(* IEC 61131-3 sources: daoli-st-library/DL_Motion (part 9) *)

(* ---- FB_DL_AxisScrewPitchComp.st ---- *)
(*==============================================================================
 * 组件名称 (Component)  : FB_DL_AxisScrewPitchComp
 * 所属子库 (Sublibrary) : DL_Motion
 * 当前版本 (Version)    : 1.0.0
 * 兼容性   (Platform)   : CODESYS 3.5+ / TwinCAT 3 / 汇川 InoProShop / 施耐德 Machine Expert
 *                         仅依赖 Standard.library（TRUNC / ABS），零厂商私有库
 * 功能描述 (Function)   : 丝杠螺距误差分段前馈补偿：误差表 aErrTable[0..nSegCnt]
 *                         给出均匀分段节点（段长 fSegLenMm，表长 = 段数 + 1，
 *                         一致性校验）处螺距误差（mm），段内线性插值：
 *                           idx  = TRUNC(fPosMm ÷ fSegLenMm)，钳位 [0, nSegCnt−1]
 *                           fFrac = fPosMm ÷ fSegLenMm − idx，钳位 [0,1]
 *                           fCompValMm = aErrTable[idx]
 *                                        + fFrac × (aErrTable[idx+1] − aErrTable[idx])
 *                         位置先钳入表覆盖域 [0, nSegCnt×fSegLenMm]（越域置
 *                         信息码 ePosClamped），段索引防越界钳位（规格指定）；
 *                         非有限位置输出 0 并置信息码 ePosNonFin（规格指定）。
 * 接口     (Interface)  : 输入 fPosMm 轴当前位置 [mm]、aErrTable 分段误差表
 *                         （定长 0..16，[mm]）、nSegCnt 有效段数（域 [1,16]）、
 *                         fSegLenMm 每段长度（域 > 0）、bReset 复位；
 *                         输出 fCompValMm 前馈补偿值（叠加到位置设定侧）
 *                         [mm]、eErrCode 错误码、bError 故障标志。
 * 边界     (Boundary)   : ① **属主边界（写死）：本件只算螺距误差补偿量，不写
 *                         位置指令、不接管反向间隙补偿**；间隙补偿归
 *                         `FB_DL_AxisBacklashComp`。
 *                         ② 表长一致性：nSegCnt 有效段数对应节点 0..nSegCnt
 *                         共 nSegCnt+1 个，超出定长 17（nSegCnt > 16）或
 *                         nSegCnt < 1 → 锁存故障（表长=段数+1 一致性校验，
 *                         规格指定），冻结输出 0。
 *                         ③ 位置域钳位：fPosMm < 0 钳 0、> nSegCnt×fSegLenMm
 *                         钳上界，置信息码 ePosClamped（量值方向可饱和）。
 *                         ④ 非有限判据（R79 双判）先行于一切换算：非有限时
 *                         输出 0、信息码 ePosNonFin，不污染插值。
 *                         ⑤ 组态闸：fSegLenMm <= 0 → 锁存故障（除数前置闸，
 *                         结构性无除零），冻结输出 0，解除沿 = bReset 上升沿。
 *                         ⑥ TRUNC 取整前位置已过非有限闸与域钳位（无溢出
 *                         取整路径）。
 *                         ⑦ 零全局耦合（无 GVL / VAR_EXTERNAL / 物理地址）。
 * 分工声明 (Scope)      : 与 `FB_DL_AxisBacklashComp` 分工：反向间隙（双区滞回）
 *                         归那件、螺距分段误差（单值表）归本件；与
 *                         `FB_DL_CamTableInterp` 分工：凸轮表插值归那件。
 * 来源标签 (Source Tag) : 自研线（分段线性插值为公开数值方法 clean-room）
 * 码表     (Codes)      : 本件不占用任何全局数字码位。出口为 LREAL 补偿值 +
 *                         ENUM 错误码；数字码位待主控收口阶段统一派号。
 * 红线自检 (Redline)    : R1 ✓ 零 GVL/VAR_EXTERNAL ｜ R2 ✓ 零 %I/%Q/%M ｜ R3 ✓ 纯 IEC 61131-3
 *                         R4 ✓ 索引钳位 + 表长一致性 + 除数前置闸 + 非有限先行
 *                         ｜ R5 ✓ 声明逐行同行双语注释
 *                         R6 N/A（无 ENUM 状态机） ｜ R7 ✓ 一 R_TRIG 段 0 无条件刷新
 * 修订历史 (Revision)   : 2026-11-20  v1.0.0  R50 首版（批次 2 · 序号 7）
 * 验收向量 (Acceptance) : ① fSegLenMm=10, nSegCnt=2, aErrTable=[0.0, 0.01, 0.03]
 *                         （mm）：fPosMm=5 → 段 0 半程 → 0.0 + 0.5×0.01 =
 *                         0.005 mm；fPosMm=15 → 段 1 半程 → 0.01 + 0.5×0.02
 *                         = 0.02 mm，均 eOk；② fPosMm=25 → 钳上界 20 → 段 1
 *                         终点 → 0.03 mm，ePosClamped；③ nSegCnt=0 → 锁存
 *                         eCfgBad，输出 0；④ fPosMm=NaN → 输出 0，
 *                         ePosNonFin。
 *==============================================================================*)

(*-----------------------------------------------------------------------------
 * 枚举: E_DL_SpcErr（错误码；信息级不置 bError，故障级恒伴 bError=TRUE）
 *----------------------------------------------------------------------------*)
TYPE E_DL_SpcErr :
(
    eOk         := 0,   // 正常 / Normal
    eCfgBad     := 1,   // 故障级：段数/段长组态非法（表长=段数+1 破坏） / Fault: segment config illegal
    ePosClamped := 2,   // 信息级：位置越表域已钳位 / Info: position clamped into table domain
    ePosNonFin  := 3    // 信息级：位置非有限，输出 0 / Info: position non-finite, output zero
);
END_TYPE

FUNCTION_BLOCK FB_DL_AxisScrewPitchComp
VAR_INPUT
    fPosMm    : LREAL := 0.0;                  // 轴当前位置 [mm] / Axis present position [mm]
    aErrTable : ARRAY[0..16] OF LREAL;         // 分段误差表（节点 0..nSegCnt） [mm] / Segmented error table [mm]
    nSegCnt   : UDINT := 8;                    // 有效段数（表长 = 段数+1），域 [1,16] [段] / Valid segment count
    fSegLenMm : LREAL := 10.0;                 // 每段长度，域 > 0 [mm] / Segment length [mm]
    bReset    : BOOL := FALSE;                 // 复位，上升沿清组态故障锁存 [-] / Reset, rising edge clears cfg latch
END_VAR
VAR_OUTPUT
    fCompValMm : LREAL;                        // 前馈补偿值（叠加位置设定侧） [mm] / Feedforward compensation [mm]
    eErrCode   : E_DL_SpcErr;                  // 错误码出口 / Error code outlet
    bError     : BOOL;                         // 故障标志（组态锁存） [-] / Error flag, latched
END_VAR
VAR
    _nIdx     : DINT;                          // 段索引（钳位后，域 [0, nSegCnt−1]） [-] / Clamped segment index
    _fScaled  : LREAL;                         // 位置按段长标度值（无量纲段数） [段] / Position scaled by segment length
    _fFrac    : LREAL;                         // 段内分数（钳位 [0,1]） [-] / In-segment fraction
    _fPosUse  : LREAL;                         // 钳入表域后的位置 [mm] / Position clamped into domain
    _fPosMax  : LREAL;                         // 表覆盖域上界 = nSegCnt×fSegLenMm [mm] / Table domain ceiling
    _bNonFin  : BOOL;                          // 位置非有限当拍量 [-] / Position non-finite this scan
    _bClamped : BOOL;                          // 本拍发生位置钳位 [-] / Position clamped this scan
    _bCfgBad  : BOOL;                          // 组态非法当拍量 [-] / Illegal configuration this scan
    _bErrLatch: BOOL;                          // 组态故障锁存位（解除沿 = bReset 上升沿） / Latched config fault
    rtReset   : R_TRIG;                        // 复位沿实例，段 0 无条件调用 / Reset edge instance
END_VAR
VAR CONSTANT
    DL_SPC_NMAX  : DINT := 16;                 // 段数上限（表定长 0..16 共 17 节点） [段] / Segment count ceiling
    DL_SPC_NMIN  : DINT := 1;                  // 段数下限 [段] / Segment count floor
    DL_SPC_ZERO  : LREAL := 0.0;               // 域下界与判零基准 [mm] / Domain floor and zero base
    DL_SPC_ONE   : LREAL := 1.0;               // 分数钳位上界 [-] / Fraction ceiling
END_VAR

(* —— 段 0：非有限判 + 组态闸 + 沿刷新 —— *)
_bNonFin := (fPosMm <> fPosMm) OR ((fPosMm - fPosMm) <> DL_SPC_ZERO);   // 位置非有限（R79 双判） / Position non-finite
_bCfgBad := (fSegLenMm <= DL_SPC_ZERO);        // 段长域闸（除数前置） / Segment length gate
IF (UDINT_TO_DINT(nSegCnt) < DL_SPC_NMIN) OR (UDINT_TO_DINT(nSegCnt) > DL_SPC_NMAX) THEN
    _bCfgBad := TRUE;                          // 表长=段数+1 一致性破坏（规格②） / Table length consistency violated
END_IF
rtReset(CLK := bReset);                        // 复位沿，每拍必调 / Reset edge, every scan

(* —— 段 1：复位沿与组态锁存 —— *)
IF rtReset.Q THEN
    _bErrLatch := FALSE;                       // 清组态锁存（R188 声明：解除沿 = bReset 上升沿） / Clear cfg latch
END_IF
IF _bCfgBad AND (NOT _bErrLatch) THEN
    _bErrLatch := TRUE;                        // 锁存 / Latch
END_IF

(* —— 段 2：位置域钳位（故障期跳过；非有限跳过） —— *)
_bClamped := FALSE;                            // 钳位量预清 / Clamp preset
_fPosUse := DL_SPC_ZERO;                       // 安全侧起步 0 / Safe-side start zero
_fPosMax := UDINT_TO_LREAL(nSegCnt) * fSegLenMm;   // 表域上界 [mm] / Domain ceiling
IF (NOT _bErrLatch) AND (NOT _bNonFin) THEN
    _fPosUse := fPosMm;                        // 位置工作副本 / Position working copy
    IF _fPosUse < DL_SPC_ZERO THEN
        _fPosUse := DL_SPC_ZERO;               // 下越域钳 0 / Clamp low to zero
        _bClamped := TRUE;                     // 记钳位 / Mark clamp
    ELSIF _fPosUse > _fPosMax THEN
        _fPosUse := _fPosMax;                  // 上越域钳上界 / Clamp high to ceiling
        _bClamped := TRUE;                     // 记钳位 / Mark clamp
    END_IF
END_IF

(* —— 段 3：分段线性插值（索引与分数双重钳位，防越界） —— *)
IF (NOT _bErrLatch) AND (NOT _bNonFin) THEN
    _fScaled := _fPosUse / fSegLenMm;          // 标度值（除数已过闸，结构性无除零） / Scaled value
    _nIdx := LREAL_TO_DINT(TRUNC(_fScaled));   // 段索引取整（域已钳，无溢出） / Segment index by TRUNC
    IF _nIdx > (UDINT_TO_DINT(nSegCnt) - 1) THEN
        _nIdx := UDINT_TO_DINT(nSegCnt) - 1;   // 索引上钳（规格：防越界钳位） / Clamp index high
    END_IF
    IF _nIdx < 0 THEN
        _nIdx := 0;                            // 索引下钳 / Clamp index low
    END_IF
    _fFrac := _fScaled - DINT_TO_LREAL(_nIdx);   // 段内分数（索引升位实数化） / In-segment fraction
    IF _fFrac < DL_SPC_ZERO THEN
        _fFrac := DL_SPC_ZERO;                 // 分数下钳 / Clamp fraction low
    END_IF
    IF _fFrac > DL_SPC_ONE THEN
        _fFrac := DL_SPC_ONE;                  // 分数上钳 / Clamp fraction high
    END_IF
    fCompValMm := aErrTable[_nIdx] + _fFrac * (aErrTable[_nIdx + 1] - aErrTable[_nIdx]);   // 段内线性插值（_nIdx+1 <= nSegCnt 表内） / Linear interpolation
ELSE
    fCompValMm := DL_SPC_ZERO;                 // 故障/非有限安全侧输出 0（规格④） / Safe-side zero output
END_IF

(* —— 段 4：出口单点映射（错误码归约，R191） —— *)
IF _bErrLatch THEN
    bError := TRUE;                            // 故障标志（R45 配对） / Error flag
    eErrCode := E_DL_SpcErr.eCfgBad;           // 故障级码 / Fault code
ELSE
    bError := FALSE;                           // 无故障级条件 / No fault
    IF _bNonFin THEN
        eErrCode := E_DL_SpcErr.ePosNonFin;    // 信息级：非有限口径 / Info: non-finite
    ELSIF _bClamped THEN
        eErrCode := E_DL_SpcErr.ePosClamped;   // 信息级：越域钳位口径 / Info: clamped
    ELSE
        eErrCode := E_DL_SpcErr.eOk;           // 正常 / Normal
    END_IF
END_IF

END_FUNCTION_BLOCK

(* ---- FB_DL_AxisSoftLimitGuard.st ---- *)
(*
    FB_DL_AxisSoftLimitGuard —— 轴软限位守卫（位置 + 速度前馈预判减速请求）
    ------------------------------------------------------------------
    组件名称  : FB_DL_AxisSoftLimitGuard
    分类      : DL_Motion / LimitGuard
    前缀      : FB_DL_
    版本      : 1.0.0
    溯源      : 借鉴点 —— 运动控制领域「软限位 + 提前减速（预判停距）」的通行语义：
                仅用位置比较只能撞限位后才发现（已超程），故必须用当前速度按
                允许减速度反算停距，把「当前位置 + 本周期位移 + 停距」作为预判
                可达位置，与限位比较后提前发出减速请求；越限后锁存并禁止该方向
                运动（方向互锁）。该语义与 PLCopen Motion Control 公开规范中
                「软限位监视 / 方向禁止」的功能描述一致。
                clean-room 声明 —— 零代码行复制；本件不含任何厂商运动指令
                （不调用 MC_* 功能块、不使用任何厂商专有数据类型），停距预判、
                方向互锁、闸门、码位与双语文档全部自有。
                许可证 —— 本件 MIT；来源标签 s7motion 仅指该语义在公开厂商文档
                中的功能描述，文档不属代码，无许可继承。
    平台      : 纯 IEC 61131-3，CODESYS 3.5 / TwinCAT 3 / InoProShop / Machine Expert 通用
    作者      : 道莅代码库 · PLC编程专家（R70 构建轮 · 批 3 · N8）
    ------------------------------------------------------------------
    功能说明  : 预判模型（逐项写清，便于现场复核）：
                  fSpan := ABS(fVel) * fScanSec               本周期位移（速度前馈项，[mm]）
                  fStop := fVel * fVel / (2 * fDecel)         停距（等减速度制动距离，[mm]）
                  fPred := fPos + fVel * fScanSec + 符号(fVel) * fStop   预判可达位置 [mm]
                判据：
                  正向减速请求 bDecelPos := fVel > 0 且 fPred > (fPosMax - fMargin)
                  负向减速请求 bDecelNeg := fVel < 0 且 fPred < (fPosMin + fMargin)
                  正向禁止 bInhibitPos := 越限锁存 或 fPos >= fPosMax
                  负向禁止 bInhibitNeg := 越限锁存 或 fPos <= fPosMin
                除法面（唯一除法）：除子为 (2 * fDecel)，进入除法前经**两道结构闸**
                校验 fDecel > 0 与 (2 * fDecel) > 0，两者同时成立才落除法；
                闸不成立时整个预判段被跳过（不落除法、不发减速请求、不写
                fPredPos），并由组态闸在段 4 置 0501 锁存。
                其余算式一律用乘加（余量比较改写为 fMargin * 2 >= 行程），
                故本件全部代码中只有一个除法点。
                越限锁存：fPos 越过任一限位即锁存 0503，bReset 上升沿解除；
                锁存期内两个禁止方向位**恒为 TRUE**（双方向全禁，因为越限后
                任何方向都可能加剧超程，需人工确认后复位）。
    错误码    : 16#0002_0501 组态非法（限位反置 / 减速度非正 / 回退余量为负 / 非有限），锁存 —— 故障级
                16#0002_0502 位置或速度非有限，锁存 —— 故障级
                16#0002_0503 越限（位置越过软限位），锁存 —— 故障级
    码位总账  : 0501 / 0502 / 0503 用（均故障级）；无信息级码（减速请求与禁止位已可观测）
    状态机    : N/A —— 无顺序相（逐拍组合判据 + 越限锁存），无 ENUM / CASE
    边界与披露: 一 组态闸（R272 逐项点名）：fPosMax > fPosMin；fDecel > 0；
                   fMargin >= 0 且 fMargin < (fPosMax - fPosMin) / 2（余量不得吞没
                   整个行程）；fScanSec > 0；上述量与 fPos / fVel 全部纳入
                   NaN 自反判 + Inf 差值自反判 + 幅值 1E9 上界筛查；
                二 定时器 / 沿实例：仅 _rtReset 一个沿实例，在段 2 无条件调用；
                   本件不含 TON / TOF / TP，故无定时器跳过风险；
                三 出口语义（R191）：bDecelPos / bDecelNeg 为**逐拍重算**的请求位，
                   bInhibitPos / bInhibitNeg 为组合位（越限锁存 或 位置到限），
                   bBeyond 为越限锁存镜像；三者名实同源、无混用；
                四 失能（bEn = FALSE）：减速请求清零、禁止位**保持有效**
                   （安全方向：失能不得放开方向禁止），bBusy 清零，锁存位不被清除；
                五 本件不做任何运动指令下发，只输出布尔许可 / 请求位，由上层
                   运动层转换为 MC_Halt / 减速倍率等动作 —— 保持硬件与厂商无关；
                六 零全局变量、零 VAR_EXTERNAL、零物理地址、零数组下标。
    修订记录  : 2026-11-22 v1.0.0 首次入库（R70 构建轮 · 批 3 · N8）
*)
FUNCTION_BLOCK FB_DL_AxisSoftLimitGuard
VAR_INPUT
    bEn       : BOOL := TRUE;              (* 使能，[标志] / the enable *)
    bReset    : BOOL := FALSE;             (* 越限复位（上升沿有效），[标志] / the overrun reset, rising edge *)
    fPos      : LREAL := 0.0;              (* 轴当前位置（编码器反馈），[mm] / the axis position feedback *)
    fVel      : LREAL := 0.0;              (* 轴当前速度（反馈或指令前馈），[mm/s] / the axis velocity *)
    fPosMax   : LREAL := 1000.0;           (* 正向软限位，[mm]，须 > fPosMin / the positive soft limit *)
    fPosMin   : LREAL := 0.0;              (* 负向软限位，[mm]，须 < fPosMax / the negative soft limit *)
    fDecel    : LREAL := 1000.0;           (* 允许减速度幅值，[mm/s^2]，须 > 0 / the allowed deceleration magnitude *)
    fScanSec  : LREAL := 0.004;            (* 任务周期折算秒数，[s]，须 > 0 / the task period in seconds *)
    fMargin   : LREAL := 20.0;             (* 提前减速余量，[mm]，须 >= 0 / the early deceleration margin *)
END_VAR
VAR_OUTPUT
    bDecelPos   : BOOL;                    (* 正向减速请求，[标志] / the positive direction deceleration request *)
    bDecelNeg   : BOOL;                    (* 负向减速请求，[标志] / the negative direction deceleration request *)
    bInhibitPos : BOOL;                    (* 正向运动禁止，[标志] / the positive direction inhibited *)
    bInhibitNeg : BOOL;                    (* 负向运动禁止，[标志] / the negative direction inhibited *)
    bBeyond     : BOOL;                    (* 越限锁存镜像，[标志] / the overrun latch image *)
    fPredPos    : LREAL;                   (* 预判可达位置（供诊断），[mm] / the predicted reachable position *)
    bBusy       : BOOL;                    (* 减速请求有效（占用中），[标志] / a deceleration request is active *)
    bValid      : BOOL;                    (* 出口可信（无锁存故障），[标志] / the outlets are trustworthy *)
    bError      : BOOL;                    (* 故障标志，锁存故障时为 TRUE / the fault flag, raised while latched *)
    nErrCode    : UDINT;                   (* 错误码，0 = 正常，锁存回放 / the error id, 0 = ok, replayed *)
END_VAR
VAR
    _rtReset    : R_TRIG;                  (* 复位上升沿实例（无条件调用）/ the reset rising edge instance *)
    _bFault     : BOOL;                    (* 组态 / 输入故障锁存位 / the configuration and input fault latch *)
    _bBeyond    : BOOL;                    (* 越限保持量，仅 bReset 上升沿解除 / the overrun hold *)
    _nCodeLatch : UDINT;                   (* 故障锁存码（0501 / 0502 / 0503）/ the fault code latch *)
    _bCfgBad    : BOOL;                    (* 组态非法标志（逐拍重算）/ the configuration fault flag *)
    _bInBad     : BOOL;                    (* 位置或速度非有限标志（逐拍重算）/ the input fault flag *)
    _fSpan      : LREAL;                   (* 本周期位移，[mm] / the travel within one period *)
    _fStop      : LREAL;                   (* 制动停距，[mm] / the braking distance *)
    _fPred      : LREAL;                   (* 预判可达位置（内部），[mm] / the predicted reachable position, internal *)
    _fSign      : LREAL;                   (* 速度符号的实数形式（1.0 / 0.0 / -1.0），[无量纲] / the velocity sign as a real *)
END_VAR
VAR CONSTANT
    DL_ASG_FMAX : LREAL := 1.0E9;          (* 非有限筛查幅值上限，[工程单位] / the finiteness screening cap *)
END_VAR

// 段 1｜出口预置（R256 统一出口预置）/ segment 1, preset every outlet
bDecelPos   := FALSE;                      // 正向减速请求预清零 / preset the positive request false
bDecelNeg   := FALSE;                      // 负向减速请求预清零 / preset the negative request false
bInhibitPos := FALSE;                      // 正向禁止预清零（段 7 按安全方向重算）/ preset the positive inhibit false
bInhibitNeg := FALSE;                      // 负向禁止预清零 / preset the negative inhibit false
bBeyond     := FALSE;                      // 越限镜像预清零 / preset the overrun image false
fPredPos    := 0.0;                        // 预判位置预置零 / preset the predicted position
bBusy       := FALSE;                      // 忙碌标志预清零 / preset the busy flag false
bValid      := FALSE;                      // 可用标志预置假，健康路径再置真 / preset valid false
bError      := FALSE;                      // 故障标志预清零 / preset the error flag false
nErrCode    := 0;                          // 错误码预置无错 / preset the code to zero
_fSign      := 0.0;                        // 速度符号预置零 / preset the sign to zero

// 段 2｜沿实例无条件调用（规则 ⑦，本件无 TON / TOF / TP）/ segment 2, the reset edge instance
_rtReset(CLK := bReset);                   // 复位沿，每周期无条件刷新 / the reset edge, refreshed every scan

// 段 3｜越限解除：唯一可到达的清除边（R188）/ segment 3, the only overrun release edge
IF _rtReset.Q THEN                         // 复位上升沿 / the reset rising edge
    _bBeyond := FALSE;                     // 解除越限保持 / release the overrun hold
    IF _nCodeLatch = 16#0002_0503 THEN     // 锁存码为越限时才清码（组态 / 输入码保持到修复）/ clear the code only when it was the overrun
        _nCodeLatch := 0;                  // 清锁存码 / clear the latched code
    END_IF
END_IF

// 段 4｜组态守卫（R272 逐项点名）/ segment 4, the configuration guard
_bCfgBad := (fPosMax <= fPosMin)                                     // 限位反置或重合 / the limits reversed or coincident
         OR (fDecel <= 0.0)                                          // 减速度非正（除子域非法）/ a non positive deceleration
         OR (fScanSec <= 0.0)                                        // 任务周期非正 / a non positive task period
         OR (fMargin < 0.0)                                          // 余量为负 / a negative margin
         OR (fMargin * 2.0 >= (fPosMax - fPosMin))                   // 余量吞没行程（改用乘 2，本式不落除法）/ the margin swallows the stroke, no division here
         OR (fPosMax <> fPosMax) OR ((fPosMax - fPosMax) <> 0.0) OR (ABS(fPosMax) > DL_ASG_FMAX)
         OR (fPosMin <> fPosMin) OR ((fPosMin - fPosMin) <> 0.0) OR (ABS(fPosMin) > DL_ASG_FMAX)
         OR (fDecel <> fDecel) OR ((fDecel - fDecel) <> 0.0) OR (ABS(fDecel) > DL_ASG_FMAX)
         OR (fScanSec <> fScanSec) OR ((fScanSec - fScanSec) <> 0.0) OR (ABS(fScanSec) > DL_ASG_FMAX)
         OR (fMargin <> fMargin) OR ((fMargin - fMargin) <> 0.0) OR (ABS(fMargin) > DL_ASG_FMAX);

// 段 5｜输入守卫：位置与速度非有限 / segment 5, the position and velocity guard
_bInBad := (fPos <> fPos) OR ((fPos - fPos) <> 0.0) OR (ABS(fPos) > (DL_ASG_FMAX * 10.0))
        OR (fVel <> fVel) OR ((fVel - fVel) <> 0.0) OR (ABS(fVel) > (DL_ASG_FMAX * 10.0));

// 段 6｜首次成因锁存（故障期不重推断，R189）/ segment 6, the first cause latch
IF NOT _bFault THEN                        // 未锁存才登记 / register only while healthy
    IF _bCfgBad THEN                       // 组态非法优先 / the configuration first
        _bFault     := TRUE;               // 置锁存 / latch it
        _nCodeLatch := 16#0002_0501;       // 故障级：组态非法 / fault level: an illegal configuration
    ELSIF _bInBad THEN                     // 输入非有限 / an input is non finite
        _bFault     := TRUE;               // 置锁存 / latch it
        _nCodeLatch := 16#0002_0502;       // 故障级：输入非有限 / fault level: an input is non finite
    END_IF
END_IF

// 段 7｜越限判定与方向禁止（安全方向：越限后双向全禁）/ segment 7, the overrun verdict and the direction inhibits
IF bEn AND NOT _bFault THEN                // 使能与无故障才判越限 / judge the overrun only while enabled and healthy
    IF (fPos > fPosMax) OR (fPos < fPosMin) THEN   // 位置越过任一软限位 / the position passed a soft limit
        IF NOT _bBeyond THEN               // 首次越限才登记码（不重推断）/ register the code once
            _bBeyond    := TRUE;           // 置越限保持 / hold the overrun
            _nCodeLatch := 16#0002_0503;   // 故障级：越限 / fault level: an overrun
        END_IF
    END_IF
    bInhibitPos := _bBeyond OR (fPos >= fPosMax);  // 正向禁止：越限锁存 或 位置到正限 / the positive inhibit
    bInhibitNeg := _bBeyond OR (fPos <= fPosMin);  // 负向禁止：越限锁存 或 位置到负限 / the negative inhibit
ELSE                                       // 失能或故障：禁止位保持安全侧（不放开）/ disabled or faulted, keep the inhibits safe
    bInhibitPos := TRUE;                   // 正向保持禁止 / keep the positive direction inhibited
    bInhibitNeg := TRUE;                   // 负向保持禁止 / keep the negative direction inhibited
END_IF

// 段 8｜预判停距与减速请求（唯一除法，除子先经结构闸）/ segment 8, the predictive request
IF bEn AND NOT _bFault AND NOT _bBeyond THEN   // 健康且未越限才做预判 / predict only while healthy and inside the limits
    IF fDecel > 0.0 THEN                       // 结构闸一：减速度为正 / gate one, the deceleration is positive
        IF (2.0 * fDecel) > 0.0 THEN           // 结构闸二：除子为正（禁除零，规则 ④）/ gate two, the divisor is positive
            _fSpan := ABS(fVel) * fScanSec;    // 本周期位移（速度前馈项）/ the travel within one period
            _fStop := (fVel * fVel) / (2.0 * fDecel); // 制动停距（唯一除法）/ the braking distance, the only division
            IF fVel > 0.0 THEN                 // 正向运动 / moving in the positive direction
                _fSign := 1.0;                 // 符号为正 / the sign is positive
            ELSIF fVel < 0.0 THEN              // 负向运动 / moving in the negative direction
                _fSign := -1.0;                // 符号为负 / the sign is negative
            ELSE                               // 静止 / at standstill
                _fSign := 0.0;                 // 符号为零（停距不计方向）/ the sign is zero
            END_IF
            _fPred := fPos + (fVel * fScanSec) + (_fSign * _fStop); // 预判可达位置 / the predicted reachable position
            fPredPos := _fPred;                // 预判位置出口（诊断用）/ the predicted position outlet
            bDecelPos := (fVel > 0.0) AND (_fPred > (fPosMax - fMargin));  // 正向提前减速请求 / the positive early request
            bDecelNeg := (fVel < 0.0) AND (_fPred < (fPosMin + fMargin));  // 负向提前减速请求 / the negative early request
        END_IF
    END_IF
END_IF

// 段 9｜出口映射（名实双出口同源，R191）/ segment 9, the outlet mapping
bBeyond  := _bBeyond;                      // 越限镜像 = 保持量 / the overrun image mirrors the hold
bBusy    := bDecelPos OR bDecelNeg;        // 减速请求有效即占用 / a request is active
bError   := _bFault OR _bBeyond;           // 故障标志 = 锁存故障 或 越限 / the fault flag, the latch or the overrun
bValid   := bEn AND NOT bError;            // 出口可信条件 / the outlets are trustworthy
IF _bBeyond THEN                           // 越限优先归因 / the overrun takes precedence
    nErrCode := 16#0002_0503;              // 故障级：越限 / fault level: an overrun
ELSE                                       // 非越限 / no overrun
    nErrCode := _nCodeLatch;               // 回放锁存码 / replay the latched code
END_IF
END_FUNCTION_BLOCK

(* ---- FB_DL_AxisSoftLimitPredict.st ---- *)
(*
  Name        : FB_DL_AxisSoftLimitPredict
  Category    : DL_Motion
  Version     : 1.0.0
  Purpose     : 软限位超程预测：按当前速度与最大减速度预算停车距离 s = v²/(2a)，与到限位余量比较，提前发出减速请求（预测式，非反应式拦截）；/ Predict soft-limit overtravel: budget the stopping distance s = v^2/(2a) from current velocity and maximum deceleration, compare with the remaining margin and raise a deceleration request in advance
  溯源        : 借 t2-4-s7-motion 的分类/参数域组织，clean-room 实现
  Boundary    : ① 组态闸：最大减速度 <= eps / 余量 <= 0 / 上限须大于下限 / 扫描周期 <= 0 → 锁存故障；
                ② 除子闸：2a 在组态闸后使用（a > eps 已保证）；v² 为乘性无除法；
                ③ 仅对「朝限位运动」的方向预测：速度为 0 时不请求减速（无预测语义）；
                ④ 输出为「请求」，不直接写速度/位置（属主边界：执行由运动控制层完成）；
                ⑤ 所有比较用容差或直比，禁浮点等值比较。
*)
TYPE E_DL_AslpState :
(
    eIdle  := 0,                             (* 未使能 / Disabled *)
    ePred  := 10,                            (* 预测运行 / Predicting *)
    eFault := 90                             (* 故障锁存相 / Fault latched *)
);
END_TYPE

TYPE E_DL_AslpCause :
(
    eNone       := 0,                        (* 无故障成因 / No cause *)
    eCfgIllegal := 1,                        (* 组态非法：减速度/余量/限位越域 / Illegal config *)
    ePhaseBad   := 2                         (* 非法相位兜底 / Illegal phase fallback *)
);
END_TYPE

FUNCTION_BLOCK FB_DL_AxisSoftLimitPredict
VAR_INPUT
    fPosNow   : REAL := 0.0;                 (* 当前实际位置 [mm] / Current position *)
    fVelNow   : REAL := 0.0;                 (* 当前速度（带符号）[mm/s] / Current velocity, signed *)
    fDecMax   : REAL := 5000.0;              (* 最大可用减速度，域 > 0 [mm/s²] / Maximum deceleration, > 0 *)
    fLimPos   : REAL := 1000.0;              (* 正向软限位 [mm] / Positive soft limit *)
    fLimNeg   : REAL := -1000.0;             (* 负向软限位 [mm] / Negative soft limit *)
    fMargin   : REAL := 5.0;                 (* 提前量（在停车距离上附加），域 >= 0 [mm] / Lead margin, >= 0 *)
    bEnable   : BOOL := TRUE;                (* 预测使能 [-] / Enable *)
    bReset    : BOOL := FALSE;               (* 复位命令，上升沿清输出与故障 [-] / Reset command *)
END_VAR
VAR_OUTPUT
    fStopDist : REAL;                        (* 停车距离预算 v²/(2a) [mm] / Budgeted stopping distance *)
    fDistPos  : REAL;                        (* 到正向限位的余量 [mm] / Remaining distance to positive limit *)
    fDistNeg  : REAL;                        (* 到负向限位的余量 [mm] / Remaining distance to negative limit *)
    bDecelReq : BOOL;                        (* 减速请求（预算 + 余量 >= 可用余量）[-] / Deceleration request *)
    bOvershoot: BOOL;                        (* 已判定越界（余量 <= 提前量）[-] / Already out of margin *)
    nDir      : INT;                         (* 运动方向：+1 正 / -1 负 / 0 停 [-] / Motion direction *)
    eState    : E_DL_AslpState;              (* 状态出口 / State outlet *)
    eCause    : E_DL_AslpCause;              (* 故障成因出口（R190 归因唯一） / Fault cause outlet *)
    bError    : BOOL;                        (* 故障锁存标志 [-] / Fault latch flag *)
END_VAR
VAR
    _eState  : E_DL_AslpState := E_DL_AslpState.eIdle;   (* 内部相位（CASE 唯一写入目标） / Internal phase *)
    _eCause  : E_DL_AslpCause := E_DL_AslpCause.eNone;   (* 故障成因锁存量 / Latched cause *)
    rtReset  : R_TRIG;                       (* 复位沿实例，段 0 无条件调用 / Reset edge instance *)
    _bFault  : BOOL;                         (* 故障锁存位 / Latched fault bit *)
    _bCfgBad : BOOL;                         (* 组态非法当拍量 / Illegal config this scan *)
    _bFinite : BOOL;                         (* 输入有限性当拍量 / Input finiteness *)
    _fStop   : REAL;                         (* 停车距离中间量 [mm] / Stopping distance intermediate *)
    _fNeed   : REAL;                         (* 预算 + 提前量（总需距）[mm] / Required distance *)
    _fAbsVel : REAL;                         (* 速度绝对値（距离预算用）[mm/s] / Absolute velocity *)
    _nDir    : INT;                          (* 方向判定中间量 [-] / Direction intermediate *)
    _fZero   : REAL;                         (* 实数零常量 [-] / Real zero constant *)
END_VAR
VAR CONSTANT
    DL_ASLP_EPS : REAL := 1.0E-6;            (* 判零容差（速度/减速度）[mm/s] / Epsilon *)
    DL_ASLP_TWO : REAL := 2.0;               (* 停车距离公式常量 2 [-] / Formula constant *)
    DL_ASLP_DIRP: INT  := 1;                 (* 正方向编码 [-] / Positive direction code *)
    DL_ASLP_DIRN: INT  := -1;                (* 负方向编码 [-] / Negative direction code *)
    DL_ASLP_DIR0: INT  := 0;                 (* 静止编码 [-] / Standstill code *)
END_VAR

(* —— 段 0：当拍判据派生 + 实例无条件刷新（R228A） —— *)
_bCfgBad := (fDecMax <= DL_ASLP_EPS)                                           (* 减速度正域闸（除零前置） / Deceleration gate *)
            OR (fMargin < 0.0)                                                 (* 提前量非负闸 / Margin gate *)
            OR ((fLimPos - fLimNeg) <= DL_ASLP_EPS);                           (* 限位区间正域闸 / Limit span gate *)
rtReset(CLK := bReset);                                                        (* 复位沿每拍必调 / Reset edge every scan *)
_bFinite := (fPosNow = fPosNow) AND (fVelNow = fVelNow)                        (* NaN 自反闸 / NaN reflex gates *)
            AND ((fPosNow - fPosNow) = (fPosNow - fPosNow))                    (* 位置 Inf 闸 / Position Inf gate *)
            AND ((fVelNow - fVelNow) = (fVelNow - fVelNow));                   (* 速度 Inf 闸 / Velocity Inf gate *)
_fZero := 0.0;                                                                 (* 零常量装载 / Zero constant load *)

(* —— 段 1：单拍量预清零（R107） —— *)
bDecelReq := FALSE;                                                            (* 减速请求预清 / Request preset *)
bOvershoot := FALSE;                                                           (* 越界判据预清 / Overshoot preset *)
nDir := DL_ASLP_DIR0;                                                          (* 方向出口预清为静止 / Direction preset *)
fStopDist := 0.0;                                                              (* 停车距离预清 / Stop distance preset *)

(* —— 段 2：复位沿处理（作用域：清故障 + 清输出 + 迁 eIdle，R283 逐项声明） —— *)
IF rtReset.Q THEN
    _bFault := FALSE;                                                          (* 清故障锁存 / Clear fault *)
    _eCause := E_DL_AslpCause.eNone;                                           (* 清成因 / Clear cause *)
    fStopDist := 0.0;                                                          (* 清距离预算出口 / Clear budget outlet *)
    fDistPos := 0.0;                                                           (* 清正向余量出口 / Clear positive margin *)
    fDistNeg := 0.0;                                                           (* 清负向余量出口 / Clear negative margin *)
    bDecelReq := FALSE;                                                        (* 清减速请求 / Clear request *)
    bOvershoot := FALSE;                                                       (* 清越界判据 / Clear overshoot *)
    nDir := DL_ASLP_DIR0;                                                      (* 方向回静止 / Direction to standstill *)
    _eState := E_DL_AslpState.eIdle;                                           (* 迁未使能相 / Back to idle *)
END_IF

(* —— 段 3：组态故障锁存（锁存至复位沿，R189） —— *)
IF _bCfgBad AND NOT _bFault THEN
    _bFault := TRUE;                                                           (* 锁存故障位 / Latch fault *)
    _eCause := E_DL_AslpCause.eCfgIllegal;                                     (* 成因：组态非法 / Cause: illegal config *)
    _eState := E_DL_AslpState.eFault;                                          (* 同步迁故障相 / Migrate to fault *)
END_IF

(* —— 段 4：CASE 主状态机（ELSE 兜底迁 eFault，红线 6） —— *)
CASE _eState OF
    E_DL_AslpState.eIdle:                                                      (* 未使能：不预测 / Disabled *)
        fDistPos := fLimPos - fPosNow;                                         (* 正向余量仍实时镜像（只读观测） / Positive margin mirror *)
        fDistNeg := fPosNow - fLimNeg;                                         (* 负向余量镜像 / Negative margin mirror *)
        IF bEnable AND NOT _bFault THEN
            _eState := E_DL_AslpState.ePred;                                   (* 使能进入预测 / Enter predicting *)
        END_IF
    E_DL_AslpState.ePred:                                                      (* 预测相：停车距离预算 + 双侧余量判据 / Predicting *)
        IF NOT bEnable THEN
            _eState := E_DL_AslpState.eIdle;                                   (* 失能回未使能 / Back to idle *)
        ELSIF _bFinite THEN
            fDistPos := fLimPos - fPosNow;                                     (* 到正向限位余量（可负 = 已越界）[mm] / Margin to positive limit *)
            fDistNeg := fPosNow - fLimNeg;                                     (* 到负向限位余量 [mm] / Margin to negative limit *)
            IF fVelNow > DL_ASLP_EPS THEN
                _nDir := DL_ASLP_DIRP;                                         (* 正方向运动 / Positive motion *)
            ELSIF fVelNow < (-DL_ASLP_EPS) THEN
                _nDir := DL_ASLP_DIRN;                                         (* 负方向运动 / Negative motion *)
            ELSE
                _nDir := DL_ASLP_DIR0;                                         (* 带内：按静止处理（不请求） / Deadband: standstill *)
            END_IF
            nDir := _nDir;                                                     (* 方向出口（名实同源，R191） / Direction outlet *)
            IF _nDir <> DL_ASLP_DIR0 THEN
                _fAbsVel := ABS(fVelNow);                                      (* 速度绝对値（距离与方向无关）[mm/s] / Absolute velocity *)
                _fStop := (_fAbsVel * _fAbsVel) / (DL_ASLP_TWO * fDecMax);     (* 停车距离 v²/(2a)：除子 2a > 0 已过闸 [mm] / Stopping distance *)
                fStopDist := _fStop;                                           (* 距离预算出口 / Budget outlet *)
                _fNeed := _fStop + fMargin;                                    (* 总需距 = 预算 + 提前量 [mm] / Required distance *)
                IF _nDir = DL_ASLP_DIRP THEN
                    IF fDistPos <= fMargin THEN
                        bOvershoot := TRUE;                                    (* 余量已不足提前量：实质越界 / Within margin: overshoot *)
                    END_IF
                    IF _fNeed >= fDistPos THEN
                        bDecelReq := TRUE;                                     (* 需距 >= 余量：提前请求减速 / Need >= margin: request *)
                    END_IF
                ELSE
                    IF fDistNeg <= fMargin THEN
                        bOvershoot := TRUE;                                    (* 负向余量不足 / Negative overshoot *)
                    END_IF
                    IF _fNeed >= fDistNeg THEN
                        bDecelReq := TRUE;                                     (* 负向请求减速 / Negative request *)
                    END_IF
                END_IF
            ELSE
                fStopDist := 0.0;                                              (* 静止：无停车距离预算 / Standstill: zero budget *)
            END_IF
        END_IF                                                                 (* 非有限输入：本拍不预测，保持输出 / Non-finite: hold *)
    E_DL_AslpState.eFault:                                                     (* 故障相：冻结保持末值，仅复位沿出 / Fault *)
        ;                                                                      (* 锁存回放（R28） / Replay from latch *)
    ELSE                                                                       (* 非法相位兜底迁安全态 / Illegal phase fallback *)
        _eState := E_DL_AslpState.eFault;                                      (* 迁故障相 / To fault *)
        _bFault := TRUE;                                                       (* 同步锁存 / Latch *)
        _eCause := E_DL_AslpCause.ePhaseBad;                                   (* 成因：非法相位 / Cause: illegal phase *)
END_CASE

(* —— 段 5：出口映射（bError/eState 同源，R191） —— *)
bError := _bFault;                                                             (* 故障标志镜像 / Fault flag mirror *)
eState := _eState;                                                             (* 状态出口 / State outlet *)
eCause := _eCause;                                                             (* 成因出口 / Cause outlet *)
END_FUNCTION_BLOCK

(* ---- FB_DL_AxisSs1StopSeq.st ---- *)
(*==============================================================================
 * 组件名称 (Component)  : FB_DL_AxisSs1StopSeq
 * 所属子库 (Sublibrary) : DL_Motion
 * 当前版本 (Version)    : 1.0.0
 * 兼容性   (Platform)   : CODESYS 3.5+ / TwinCAT 3 / 汇川 InoProShop / 施耐德 Machine Expert
 *                         仅依赖 Standard.library（TON / R_TRIG / ABS），零厂商私有库
 * 功能描述 (Function)   : SS1 类停止时序编排（IEC 60204-1 停止类别 1 的公开语义：先可控减速、
 *                         到位后再切转矩）。相序：eIdle → eDecel（发减速停止请求，监视速度降到
 *                         fZeroSpeedThr）→ eSettle（零速稳定 tSettleTime）→ eStoRequest
 *                         （输出 bStoRequest = TRUE）→ eDone。任一步超时（tDecelMax / tSettleMax）
 *                         进 eFault 并置码，**且 bStoRequest 仍置真**（安全侧：宁可切转矩也不
 *                         放任轴继续动）。
 * 安全声明 (Safety)     : **本件只做停止时序与 STO 请求位，不实现任何安全认证功能**
 *                         （ISO 13849 / IEC 62061 的认证、双通道架构、诊断覆盖率证明均不在本库
 *                         范围）。bStoRequest 是**请求**而非安全输出：真实安全转矩关断必须由
 *                         认证安全模块执行，本件输出不得直接驱动安全继电器。
 * 接口     (Interface)  : 输入 bStopReq 停止请求、fSpeed 实测速度、fZeroSpeedThr 零速阈值、
 *                         tDecelMax 减速相超时、tSettleTime 零速稳定时长、tSettleMax 稳定相超时、
 *                         bReset 复位；输出 bStoRequest STO 请求位、fSpeedAtStop 首次进零速时
 *                         的速度快照、eState / eCause / bError / nErrId。
 * 边界     (Boundary)   : ① 组态闸：fZeroSpeedThr <= 0.0、tDecelMax <= T#0S、tSettleMax <= T#0S、
 *                         tSettleTime <= T#0S、fSpeed 为 NaN → **组态非法时 bStoRequest 直接置真**
 *                         （安全侧优先于组态正确性：宁可误切转矩也不放过运动轴）；
 *                         ② 零速判据用容差式（ABS <= 阈值），禁浮点判等；
 *                         ③ TON 三枚 + R_TRIG 一枚段 0 无条件周期刷新，IN 由相位派生（R228A）；
 *                         ④ 故障相迁出唯一路径 = bReset 上升沿，迁出后回 eIdle；
 *                         ⑤ 零全局耦合（无 GVL / 无物理地址）。
 * 解除式   (Release)    : bReset 上升沿 ∧ 组态合法 ∧ 速度快照已在阈值内（ABS(fSpeed) <= fZeroSpeedThr，
 *                         当拍量，R240 范式）。自证可满足（终审两式 1）：轴停住后速度快照必入阈值，
 *                         解除式不含计时器输出，无恒假因子；轴仍转时不允许解除是设计意图
 *                         （防止带速复位把 STO 请求抹掉）。
 * 码表     (Codes)      : 16#0004_03B5 故障级：SS1 停止时序故障总码（组态非法 / 减速超时 / 稳定超时 /
 *                         非法相位），锁存至 bReset 上升沿，归因由 eCause 承载（R190 单件单总码）；
 *                         16#0004_04B5 信息级：SS1 停止序列正常完成（进 eDone 单拍）。
 *                         加码反证（R90）：完成时 bStoRequest 恒为真、eState 也为固定值，正常完成与
 *                         「一直停在 eStoRequest」在出口组合上只差相位值，而相位不是台账事件，
 *                         故立一码记录每一次成功停止行程。
 *                         码段说明：0004 段故障子带 03xx / 信息子带 04xx，本件取 03B5 / 04B5
 *                         （源码实扫该两槽为空，续接同子带已用最大值，未回填碎片孔洞）。
 * 开源溯源 (Origin)     : 道莅自研 clean-room（参考 IEC 60204-1 公开停止类别语义与
 *                         t1-6-plcopen 参数域，零代码行复制）
 * 修订历史 (Revision)   : 2026-11-19  v1.0.0  R45 首版（批次 3 · 序号 11）
 *==============================================================================*)

TYPE E_DL_Ss1State :
(
    eIdle      := 0,     // 待停止请求 / Idle, awaiting stop request
    eDecel     := 10,    // 减速相：等速度降到零速阈值 / Decelerating to zero speed
    eSettle    := 20,    // 稳定相：零速保持 tSettleTime / Settling at zero speed
    eStoRequest := 30,   // STO 请求相：bStoRequest 置真 / STO request asserted
    eDone      := 50,    // 停止完成 / Stop sequence done
    eFault     := 90     // 故障锁存相（bStoRequest 仍为真） / Fault latched, STO request still TRUE
);
END_TYPE

TYPE E_DL_Ss1Cause :
(
    eNone       := 0,    // 无故障成因 / No cause
    eCfgIllegal := 1,    // 组态非法 / Illegal configuration
    eDecelTmo   := 2,    // 减速相超时 / Decel phase timeout
    eSettleTmo  := 3,    // 稳定相超时 / Settle phase timeout
    ePhaseBad   := 4     // 非法相位兜底 / Illegal phase fallback
);
END_TYPE

FUNCTION_BLOCK FB_DL_AxisSs1StopSeq
VAR_INPUT
    bStopReq      : BOOL := FALSE;        // 停止请求（电平，撤除则回空闲） [-] / Stop request level, release returns idle
    fSpeed        : REAL := 0.0;          // 实测速度（幅值判零速，符号不参与） [mm/s] / Measured speed, sign ignored [mm/s]
    fZeroSpeedThr : REAL := 5.0;          // 零速阈值，域 > 0.0 [mm/s] / Zero-speed threshold, domain > 0.0 [mm/s]
    tDecelMax     : TIME := T#5S;         // 减速相超时，域 > T#0S [ms] / Decel phase timeout, domain > T#0S [ms]
    tSettleTime   : TIME := T#200MS;      // 零速稳定时长，域 > T#0S [ms] / Zero-speed settle duration [ms]
    tSettleMax    : TIME := T#3S;         // 稳定相超时，域 > T#0S 且 >= tSettleTime [ms] / Settle phase timeout [ms]
    bReset        : BOOL := FALSE;        // 复位命令，上升沿清故障 [-] / Reset command, rising edge clears fault
END_VAR
VAR_OUTPUT
    bStoRequest   : BOOL;                 // STO 请求位（请求不等于安全认证输出） [-] / STO request, not a certified safety output
    fSpeedAtStop  : REAL;                 // 首次进零速时的速度快照 [mm/s] / Speed snapshot at first zero-speed entry
    eState        : E_DL_Ss1State;        // 状态出口，段 6 单点映射 / State outlet
    eCause        : E_DL_Ss1Cause;        // 故障成因出口（R190 归因唯一） / Fault cause outlet
    bError        : BOOL;                 // 故障锁存标志 [-] / Fault latch flag
    nErrId        : UDINT;                // 事件码，0 = 无事件 / Event code, 0 = no event
END_VAR
VAR
    _eState       : E_DL_Ss1State := E_DL_Ss1State.eIdle;   // 内部相位（CASE 唯一写入目标） / Internal phase
    _eCause       : E_DL_Ss1Cause := E_DL_Ss1Cause.eNone;   // 故障成因锁存（锁存量） / Latched cause
    tonDecel      : TON;                  // 减速相计时，段 0 无条件调用 / Decel phase timer
    tonSettle     : TON;                  // 稳定相超时计时，段 0 无条件调用 / Settle timeout timer
    tonSettleOk   : TON;                  // 零速稳定计时，段 0 无条件调用 / Zero-speed settle timer
    rtReset       : R_TRIG;               // 复位沿实例，段 0 无条件调用 / Reset edge
    _fSpeedAtStop : REAL;                 // 速度快照（锁存量，进稳定相时锁存一次） [mm/s] / Speed snapshot, latched on settle entry
    _bSnapshotOk  : BOOL;                 // 快照已锁存标记（锁存量） [-] / Snapshot taken flag
    _bZeroSpeed   : BOOL;                 // 零速当拍量 [-] / Zero-speed verdict this scan
    _bNonFin      : BOOL;                 // 速度非有限当拍量 [-] / Non-finite speed this scan
    _bCfgBad      : BOOL;                 // 组态非法当拍量 [-] / Illegal configuration
    _bStoReq      : BOOL;                 // STO 请求内部位（由相位派生） [-] / Internal STO request, derived from phase
    _bFault       : BOOL;                 // 故障锁存位（锁存量） / Latched fault bit
    _uFault       : UDINT;                // 故障码锁存（锁存量） / Latched fault code
    _uInfo        : UDINT;                // 信息码，每拍重算 / Info code, recomputed each scan
END_VAR
VAR CONSTANT
    DL_SPEED_EPS : REAL := 1.0E-3;        // 速度判零辅助容差（阈值叠加用，防阈值给到极小值） [mm/s] / Speed epsilon added to threshold [mm/s]
END_VAR

(* —— 段 0：当拍判据派生 + 定时器与沿实例无条件周期刷新 —— *)
_bNonFin    := (fSpeed <> fSpeed) OR ((fSpeed - fSpeed) <> (fSpeed - fSpeed));      // NaN 自反 + Inf 差值自减双判（判等禁令唯一例外） / NaN and Inf detection
_bZeroSpeed := ABS(fSpeed) <= (fZeroSpeedThr + DL_SPEED_EPS);                      // 零速判据（容差式） / Zero-speed verdict, tolerance-based
_bCfgBad    := (fZeroSpeedThr <= 0.0) OR (tDecelMax <= T#0S)                        // 组态域闸（R151 全覆盖） / Config gate
               OR (tSettleMax <= T#0S) OR (tSettleTime <= T#0S)                     // 时间正域闸 / Time gates
               OR (tSettleTime > tSettleMax) OR _bNonFin;                           // 配比约束：稳定时长不得超过稳定相超时 / Ratio constraint and non-finite speed
rtReset(CLK := bReset);                                                             // 复位沿，每拍必调（R228A） / Reset edge
tonDecel(IN := (_eState = E_DL_Ss1State.eDecel), PT := tDecelMax);                  // 减速相计时（IN 由相位派生） / Decel timer
tonSettle(IN := (_eState = E_DL_Ss1State.eSettle), PT := tSettleMax);               // 稳定相超时计时 / Settle timeout timer
tonSettleOk(IN := (_eState = E_DL_Ss1State.eSettle) AND _bZeroSpeed, PT := tSettleTime);   // 零速稳定计时 / Zero-speed settle timer

(* —— 段 1：单拍量预清零（锁存量与快照量不入清单，R107） —— *)
_uInfo   := 16#0000_0000;          // 信息码每拍重算 / Info recomputed every scan
nErrId   := 16#0000_0000;          // 事件码缺省无事件 / Event code default none
bError   := FALSE;                 // 故障标志每拍预清，故障分支同拍置位（R45 配对） / Flag preset
_bStoReq := FALSE;                 // STO 请求内部位缺省假，由相位与故障分支赋值 / STO internal preset

(* —— 段 2：复位沿 + 组态域闸 —— *)
IF rtReset.Q THEN                                                        // 当拍复位沿 / current-scan reset edge
    _bFault := FALSE;                                                    // 清故障锁存位（锁存量） / Clear fault latch
    _uFault := 16#0000_0000;                                             // 清故障锁存码（锁存量） / Clear latched code
    _eCause := E_DL_Ss1Cause.eNone;                                      // 清成因（锁存量） / Clear latched cause
    _bSnapshotOk := FALSE;                                               // 快照重新武装 / Re-arm snapshot
    IF _eState = E_DL_Ss1State.eFault THEN
        _eState := E_DL_Ss1State.eIdle;                                  // 故障相迁出唯一路径 / Sole exit from fault phase
    END_IF
END_IF
IF _bCfgBad THEN                                                         // 组态域闸：安全侧直接置 STO 请求 / Config gate, STO request asserted for safety
    _uFault := 16#0004_03B5;                                             // 故障级：SS1 停止时序故障总码 / Fault-level: stop-sequence fault code
    _bFault := TRUE;
    bError  := TRUE;                                                     // 故障标志同拍置位（R45 配对） / Error flag set same scan
    _eCause := E_DL_Ss1Cause.eCfgIllegal;                                // 归因：组态非法 / Cause: illegal configuration
    _bStoReq := TRUE;                                                    // 安全侧：组态非法也切转矩 / Safety side, assert STO even on bad config
END_IF

(* —— 段 3：相位派生 STO 请求（请求相 / 完成相 / 故障相均为真） —— *)
IF (_eState = E_DL_Ss1State.eStoRequest) OR (_eState = E_DL_Ss1State.eDone)
   OR (_eState = E_DL_Ss1State.eFault) THEN
    _bStoReq := TRUE;                                                    // 请求相起保持真（停住后不撤销） / Asserted from request phase onward
END_IF

(* —— 段 4：超时判据（减速相 / 稳定相） —— *)
IF (NOT _bFault) AND tonDecel.Q THEN                                     // 减速相超时 / Decel timeout
    _uFault := 16#0004_03B5;
    _bFault := TRUE;
    bError  := TRUE;
    _eCause := E_DL_Ss1Cause.eDecelTmo;                                  // 归因：减速超时 / Cause: decel timeout
    _bStoReq := TRUE;                                                    // 安全侧：宁可切转矩也不放任继续动 / Safety side, assert STO
END_IF
IF (NOT _bFault) AND tonSettle.Q THEN                                    // 稳定相超时 / Settle timeout
    _uFault := 16#0004_03B5;
    _bFault := TRUE;
    bError  := TRUE;
    _eCause := E_DL_Ss1Cause.eSettleTmo;                                 // 归因：稳定超时 / Cause: settle timeout
    _bStoReq := TRUE;                                                    // 安全侧 / Safety side
END_IF

(* —— 段 5：故障解除式（R240 全当拍量；轴仍转时不允许解除是设计意图） —— *)
IF rtReset.Q AND (NOT _bCfgBad) AND _bZeroSpeed THEN
    _bFault := FALSE;                                                    // 清故障锁存位（锁存量） / Clear fault latch
    _uFault := 16#0000_0000;                                             // 清故障锁存码（锁存量） / Clear latched code
    _eCause := E_DL_Ss1Cause.eNone;                                      // 清成因（锁存量） / Clear latched cause
END_IF

(* —— 段 5A：故障锁存相位迁移闸 —— *)
IF _bFault AND (_eState <> E_DL_Ss1State.eFault) THEN
    _eState := E_DL_Ss1State.eFault;                                     // 锁存即入故障相 / Latch enters fault phase
END_IF

(* —— 段 6：相位机（ENUM 全成员显式标签 + ELSE 兜底，R128） —— *)
CASE _eState OF

E_DL_Ss1State.eIdle:
    IF bStopReq AND (NOT _bFault) THEN                                   // 出口 1：收到停止请求 / Stop requested
        _eState := E_DL_Ss1State.eDecel;
    ELSIF _bFault THEN                                                   // 出口 2：故障锁存 / Fault latched
        _eState := E_DL_Ss1State.eFault;
    END_IF

E_DL_Ss1State.eDecel:
    IF _bZeroSpeed THEN                                                  // 出口 1：速度已降到阈值 / Speed reached threshold
        IF NOT _bSnapshotOk THEN
            _fSpeedAtStop := fSpeed;                                     // 速度快照锁存一次（锁存量） / Latch speed snapshot once
            _bSnapshotOk := TRUE;
        END_IF
        _eState := E_DL_Ss1State.eSettle;                                // 进稳定相 / Enter settle phase
    ELSIF NOT bStopReq THEN                                              // 出口 2：撤销请求（前置消失，R98） / Request released
        _eState := E_DL_Ss1State.eIdle;
    END_IF

E_DL_Ss1State.eSettle:
    IF tonSettleOk.Q THEN                                                // 出口 1：零速稳定达标 / Zero-speed settled
        _bStoReq := TRUE;                                                // 进相同拍即置请求位（不等下一拍） / Assert request in the same scan
        _eState := E_DL_Ss1State.eStoRequest;                            // 进 STO 请求相 / Enter STO request phase
    ELSIF NOT bStopReq THEN                                              // 出口 2：撤销请求 / Request released
        _eState := E_DL_Ss1State.eIdle;
    END_IF

E_DL_Ss1State.eStoRequest:
    IF bStopReq AND _bZeroSpeed THEN                                     // 出口 1：停稳（请求位保持真） / Stopped, request stays TRUE
        _uInfo := 16#0004_04B5;                                          // 信息级：SS1 停止序列正常完成 / Info: stop sequence completed
        _eState := E_DL_Ss1State.eDone;
    ELSIF NOT bStopReq THEN                                              // 出口 2：撤销请求（前置消失，R98） / Request released
        _eState := E_DL_Ss1State.eIdle;
    END_IF

E_DL_Ss1State.eDone:
    IF NOT bStopReq THEN                                                 // 出口 1：撤销请求回空闲 / Request released returns idle
        _eState := E_DL_Ss1State.eIdle;
    ELSIF _bFault THEN                                                   // 出口 2：故障锁存 / Fault latched
        _eState := E_DL_Ss1State.eFault;
    END_IF

E_DL_Ss1State.eFault:
    ;                                                                     // 故障相：仅段 5 复位沿可迁出 / Only the reset edge leaves this phase

ELSE
    _uFault := 16#0004_03B5;                                             // 故障级：非法相位兜底（归并总码） / Illegal-phase fallback
    _bFault := TRUE;
    bError  := TRUE;
    _eCause := E_DL_Ss1Cause.ePhaseBad;                                  // 归因：非法相位 / Cause: illegal phase
    _bStoReq := TRUE;                                                    // 安全侧：非法相位同样切转矩 / Safety side on illegal phase
    _eState := E_DL_Ss1State.eFault;

END_CASE

(* —— 段 7：出口单点映射（名实同源；锁存码回放；安全侧优先） —— *)
bStoRequest  := _bStoReq OR _bFault;                                     // STO 请求 = 相位派生 ∨ 故障锁存（安全侧优先） / STO request, safety side first
fSpeedAtStop := _fSpeedAtStop;                                           // 速度快照出口（锁存量回放） / Speed snapshot outlet
IF _bFault THEN
    nErrId := _uFault;                                                   // 故障锁存码回放 / Replay latched fault code
ELSE
    nErrId := _uInfo;                                                    // 信息码 / Info code
END_IF
bError := _bFault;                                                       // 故障标志与锁存同源（名实双出口，R191） / Flag from latch
eState := _eState;                                                       // 状态出口 / State outlet
eCause := _eCause;                                                       // 成因出口 / Cause outlet

END_FUNCTION_BLOCK

(* ---- FB_DL_AxisSynchronizedStop.st ---- *)
(*
    FB_DL_AxisSynchronizedStop —— 受控同步停车
    ------------------------------------------------------------------
    分类      : DL_Motion / Motion
    前缀      : FB_DL_
    版本      : 1.0.0
    溯源      : T1-6 PLCopen Motion（只借 MC_Stop / MC_Halt 的公开「按减速度停车 +
                完成确认」语义；不实现运动核、不定义轴状态机）；停止距离解析式与
                状态映射 100% 自有；clean-room 重写，未复制任何闭源厂商源码，
                参考实现仅限 MIT/Apache 许可
    平台      : 纯 IEC 61131-3，CODESYS V3.5+ / TwinCAT 3 / InoProShop 通用
    作者      : 道莅代码库 · PLC编程专家（R18）
    ------------------------------------------------------------------
    功能说明  : 给上层运动接口生成「按固定减速度斜坡停车」的指令序列，并预估停止距离
                与停止位置；用于安全门打开、料尽、下游堵塞等需要「减速停而非自由滑行」
                的工况；本件不直接驱动伺服，零全局耦合，也不承担急停（急停由安全
                回路直连，不经本件，头注释显式声明）；
                三道闸：减速度闸（减速度为 0 或负会让「停车」永不完成，首要防御）→
                快照非有限闸 → 状态机 ELSE 兜底闸（02DA 为本件专用兜底码）；
                启动时已静止则跳过硬坡直接判完成，避免定时器空转产生假 Done。
    错误码    : 16#0004_01C9 启动时已静止（速度低于阈值），跳过斜坡直接判完成——信息级，不置故障
                16#0004_01CA 预留禁用（信息级，不得挪用）
                16#0004_02D8 减速度非法（小于 1 mm/s2），停车不可完成——故障级，转故障态
                16#0004_02D9 速度或位置快照非有限（NaN / 正负 INF）——故障级，转故障态
                16#0004_02DA 状态机落 ELSE 兜底（非法状态，一律回安全态）——用途固定，不得改作他用
    码位总账  : 16#0004_01C9 用 / 16#0004_01CA 预留 ｜ 16#0004_02D8 用 / 16#0004_02D9 用 / 16#0004_02DA 用
    状态机    : E_DL_StopState（eIdle / eRamping / eSettling / eDone / eFault），
                CASE 含 ELSE 兜底，兜底固定置 eFault、位号 99 与 02DA
    采样约定  : 三个 R_TRIG 与 fbSettle 在本体首部无条件调用；fbSettle 的 IN 引脚取上一拍
                状态判据，属正常的单拍延迟，不影响完成确认的正确性。
    修订记录  : 2026-11-16 v1.0.0 首次入库（R18）
*)

(*-----------------------------------------------------------------------------
 * 枚举: E_DL_StopState（归属本功能块，与其同文件发布）
 * 含义: 受控停车状态机离散态，步长 10 留空位，故障态取 99 排末位
 *----------------------------------------------------------------------------*)
TYPE E_DL_StopState :
(
    eIdle     := 0,    // 空闲：未收到停车请求 / Idle, no stop request received
    eRamping  := 10,   // 减速中：等待速度跌到判静止阈值以下 / Ramping, waiting for the speed to fall below the standstill threshold
    eSettling := 20,   // 稳定确认中：速度已达阈值，等待稳定窗到期 / Settling, the speed reached the threshold and the settle window is running
    eDone     := 30,   // 完成：已静止且稳定窗到期 / Done, stopped and the settle window expired
    eFault    := 99    // 故障：减速度或快照非法、被中止、或落入兜底 / Fault, illegal deceleration or snapshot, aborted, or fell into the fallback
) UINT;
END_TYPE

FUNCTION_BLOCK FB_DL_AxisSynchronizedStop
VAR_INPUT
    bEnable        : BOOL;                     // 使能，FALSE 清指令并回空闲 / enable, FALSE clears the command and returns to idle
    bExecute       : BOOL;                     // 上升沿启动停车序列 / rising edge starts the stop sequence
    bAbort         : BOOL;                     // 上升沿中止并转故障态（急停由安全回路直连，不经本件）/ rising edge aborts into the fault state, the emergency stop is hardwired elsewhere
    bReset         : BOOL;                     // 上升沿清故障回空闲 / rising edge clears the fault and returns to idle
    fActVelocity   : REAL := 0.0;              // 当前速度，由运动层注入 [mm/s] / current speed injected by the motion layer [mm/s]
    fActPosition   : REAL := 0.0;              // 当前位置，用于算停止点 [mm] / current position used for the stop point [mm]
    fDeceleration  : REAL := 500.0;            // 停车减速度 [mm/s2]，范围 1.0~1.0E5 / stop deceleration [mm/s2], range 1.0~1.0E5
    tDelayTime     : TIME := T#100MS;          // 从发出到实际减速的传动延迟 [ms]，范围 0~2000 / drive train delay from command to real deceleration [ms], range 0~2000
    fVelocityEps   : REAL := 0.5;              // 判静止的速度阈值 [mm/s]，范围 0.01~100.0 / standstill speed threshold [mm/s], range 0.01~100.0
END_VAR
VAR_OUTPUT
    bBusy         : BOOL;                      // 停车进行中 / stop in progress
    bDone         : BOOL;                      // 已完成，单周期脉冲 / completed, single-cycle pulse
    bStopped      : BOOL;                      // 已静止（速度低于阈值且稳定窗到期）/ stopped, the speed is below the threshold and the settle window expired
    fStopDistance : REAL;                      // 预估停止距离（延迟段加减速段）[mm] / estimated stop distance, delay segment plus ramp segment [mm]
    fStopPosition : REAL;                      // 预估停止位置 [mm] / estimated stop position [mm]
    uState        : UINT;                      // 状态镜像 0 空闲 / 10 减速 / 20 稳定 / 30 完成 / 99 故障，仅供 HMI / state mirror for the HMI only
    eErr          : UDINT;                     // 错误码，0=正常 / error id, 0=ok
    bError        : BOOL;                      // 故障标志，eErr 为故障级时 TRUE / error flag, TRUE on fault-level eErr
END_VAR
VAR
    fbTrigExec   : R_TRIG;                     // 启动沿检测实例，本体首部无条件刷新 / execute edge instance, refreshed unconditionally
    fbTrigAbort  : R_TRIG;                     // 中止沿检测实例，本体首部无条件刷新 / abort edge instance, refreshed unconditionally
    fbTrigReset  : R_TRIG;                     // 复位沿检测实例，本体首部无条件刷新 / reset edge instance, refreshed unconditionally
    fbSettle     : TON;                        // 稳定窗定时器，本体首部无条件刷新 / settle window timer, refreshed unconditionally
    eState       : E_DL_StopState := E_DL_StopState.eIdle; // 内部状态机步序 / internal state machine step
    fDecelEff    : REAL;                       // 生效减速度，钳位后使用 [mm/s2] / effective deceleration after clamping [mm/s2]
    fStopDistCalc: REAL;                       // 停止距离计算中间量 [mm] / stop distance intermediate [mm]
    tRampCalc    : TIME;                       // 理论减速段时长，供 HMI 排程 [ms] / theoretical ramp duration for HMI scheduling [ms]
    fAbsVel      : REAL;                       // 速度绝对值 [mm/s] / absolute speed [mm/s]
    fDelaySec    : REAL;                       // 传动延迟秒值 [s] / drive train delay in seconds [s]
    fVelEpsEff   : REAL;                       // 生效判静止阈值 [mm/s] / effective standstill threshold [mm/s]
    bNonFin      : BOOL;                       // 快照非有限判定标志 / snapshot non-finite flag
END_VAR
VAR CONSTANT
    DL_STOP_DEC_MIN   : REAL := 1.0;           // 减速度下限 [mm/s2] / deceleration lower bound [mm/s2]
    DL_STOP_DEC_MAX   : REAL := 1.0E5;         // 减速度上限，超此值钳位但不判故障（高减速度是合法急停辅助）[mm/s2] / deceleration upper bound, clamped without a fault because a high value is a legal stop aid [mm/s2]
    DL_STOP_VEL_MIN   : REAL := 0.01;          // 判静止阈值下限 [mm/s] / standstill threshold lower bound [mm/s]
    DL_STOP_VEL_MAX   : REAL := 100.0;         // 判静止阈值上限 [mm/s] / standstill threshold upper bound [mm/s]
    DL_STOP_SETTLE    : TIME := T#100MS;       // 稳定确认窗 [ms] / settle confirmation window [ms]
    DL_STOP_MS_SEC    : REAL := 1000.0;        // 毫秒转秒的除数，恒非零 [ms/s] / milliseconds to seconds divisor, never zero [ms/s]
    DL_STOP_TWO       : REAL := 2.0;           // 减速段距离式的常数二 [无量纲] / constant two of the ramp distance formula [dimensionless]
    DL_FLOAT_EPS      : REAL := 1.0E-6;        // 浮点判等容差 [mm/s] / float equality tolerance [mm/s]
    DL_STOP_INF_GUARD : REAL := 4.0E38;        // 非有限幅值判定阈值 [mm] / non-finite magnitude guard [mm]
    DL_STOP_UI_IDLE   : UINT := 0;             // 状态镜像：空闲 / state mirror, idle
    DL_STOP_UI_RAMP   : UINT := 10;            // 状态镜像：减速中 / state mirror, ramping
    DL_STOP_UI_SETTLE : UINT := 20;            // 状态镜像：稳定确认中 / state mirror, settling
    DL_STOP_UI_DONE   : UINT := 30;            // 状态镜像：完成 / state mirror, done
    DL_STOP_UI_FAULT  : UINT := 99;            // 状态镜像：故障 / state mirror, fault
    DL_STOP_ZERO      : REAL := 0.0;           // 零值常量，避免裸字面量 [无量纲] / zero constant, avoids a bare literal [dimensionless]
END_VAR

// 段 1｜边沿与定时器实例无条件周期刷新（红线：严禁放入条件分支）/ segment 1, unconditional refresh of the edges and the timer
fbTrigExec(CLK := bExecute);
fbTrigAbort(CLK := bAbort);
fbTrigReset(CLK := bReset);
fbSettle(IN := (eState = E_DL_StopState.eSettling), PT := DL_STOP_SETTLE); // IN 取上一拍状态，属正常单拍延迟 / the IN pin uses the previous cycle state, a normal one-cycle lag

// 段 2｜输出与错误状态预置 / segment 2, preset outputs and error status
bDone := FALSE;                                // 完成脉冲先清 / clear the done pulse first
eErr := 0;                                     // 预置无错误 / preset no error
bError := FALSE;                               // 预置无故障 / preset no fault

// 段 3｜使能闸：失能清指令回空闲 / segment 3, enable gate returns to idle
IF NOT bEnable THEN
    eState := E_DL_StopState.eIdle;            // 回空闲态 / back to idle
    bBusy := FALSE;                            // 清忙标志 / clear the busy flag
    bStopped := FALSE;                         // 清静止标志 / clear the stopped flag
    uState := DL_STOP_UI_IDLE;                 // 状态镜像回 0 / state mirror back to zero
    RETURN;                                    // 失能即出口 / disabled is the exit
END_IF

// 段 4｜减速度闸：0 或负会让停车永不完成，是本件首要防御 / segment 4, deceleration gate
IF fDeceleration < DL_STOP_DEC_MIN THEN
    fDecelEff := DL_STOP_DEC_MIN;              // 给安全值，避免后续除零 / use the safe value so later divisions stay legal
    eErr := 16#0004_02D8;                      // 减速度非法故障码 / illegal deceleration fault id
    bError := TRUE;                            // 置故障标志 / raise the error flag
    eState := E_DL_StopState.eFault;           // 转故障态 / enter the fault state
ELSIF fDeceleration > DL_STOP_DEC_MAX THEN
    fDecelEff := DL_STOP_DEC_MAX;              // 超上限钳位，不判故障 / clamp above the upper bound without a fault
ELSE
    fDecelEff := fDeceleration;                // 域内沿用 / use the value inside the domain
END_IF
fVelEpsEff := MIN(MAX(fVelocityEps, DL_STOP_VEL_MIN), DL_STOP_VEL_MAX); // 判静止阈值双侧钳位 / clamp the standstill threshold both sides

// 段 5｜快照非有限闸：速度或位置非法即转故障态 / segment 5, non-finite snapshot gate
bNonFin := (fActVelocity <> fActVelocity)
        OR (fActVelocity > DL_STOP_INF_GUARD) OR (fActVelocity < -DL_STOP_INF_GUARD)
        OR (fActPosition <> fActPosition)
        OR (fActPosition > DL_STOP_INF_GUARD) OR (fActPosition < -DL_STOP_INF_GUARD); // 双快照同口径检查 / both snapshots checked the same way
IF bNonFin THEN
    eErr := 16#0004_02D9;                      // 快照非有限故障码 / non-finite snapshot fault id
    bError := TRUE;                            // 置故障标志 / raise the error flag
    eState := E_DL_StopState.eFault;           // 转故障态 / enter the fault state
END_IF

// 段 6｜中止与复位沿（中止优先于复位；中止是人為合法操作，不额外置参数码）/ segment 6, abort and reset edges
IF fbTrigAbort.Q THEN
    eState := E_DL_StopState.eFault;           // 中止转故障态 / an abort enters the fault state
    bBusy := FALSE;                            // 清忙标志 / clear the busy flag
    bStopped := FALSE;                         // 清静止标志 / clear the stopped flag
END_IF
IF fbTrigReset.Q THEN
    eState := E_DL_StopState.eIdle;            // 复位回空闲 / reset returns to idle
    eErr := 0;                                 // 复位清错误码 / reset clears the error id
    bError := FALSE;                           // 复位清故障标志 / reset clears the error flag
END_IF

// 段 7｜速度绝对值与停止距离预备 / segment 7, absolute speed and stop distance preparation
fAbsVel := ABS(fActVelocity);                  // 速度绝对值 / absolute speed
fDelaySec := TIME_TO_REAL(tDelayTime) / DL_STOP_MS_SEC; // 传动延迟秒值 / drive train delay in seconds

// 段 8｜状态机主体（CASE 必含 ELSE 兜底，红线）/ segment 8, state machine body
CASE eState OF
    E_DL_StopState.eIdle :
        bBusy := FALSE;                        // 空闲不忙 / idle is not busy
        bStopped := FALSE;                     // 空闲不算静止 / idle does not count as stopped
        uState := DL_STOP_UI_IDLE;             // 状态镜像 / state mirror
        IF fbTrigExec.Q THEN
            fStopDistCalc := fAbsVel * fDelaySec
                           + (fAbsVel * fAbsVel) / (DL_STOP_TWO * fDecelEff); // 延迟段加减速段，分母已由段 4 保证非零 / delay segment plus ramp segment, the divisor passed the gate in segment four
            fStopDistance := fStopDistCalc;    // 对外发布停止距离 / publish the stop distance
            IF fActVelocity >= DL_STOP_ZERO THEN
                fStopPosition := fActPosition + fStopDistCalc; // 正向运动，停止点在当前位之前 / moving positive, the stop point lies ahead
            ELSE
                fStopPosition := fActPosition - fStopDistCalc; // 反向运动 / moving negative
            END_IF
            tRampCalc := REAL_TO_TIME(fAbsVel / fDecelEff * DL_STOP_MS_SEC); // 理论减速段时长 / theoretical ramp duration
            IF fAbsVel <= fVelEpsEff THEN
                eState := E_DL_StopState.eSettling; // 本来已停，直接进稳定确认 / already stopped, go straight to settling
                eErr := 16#0004_01C9;          // 已静止提示（信息级不置故障）/ already stopped hint, info level never raises a fault
            ELSE
                eState := E_DL_StopState.eRamping; // 需要真实减速段 / a real ramp is required
            END_IF
        END_IF
    E_DL_StopState.eRamping :
        bBusy := TRUE;                         // 减速中 / ramping
        uState := DL_STOP_UI_RAMP;             // 状态镜像 / state mirror
        IF fAbsVel <= fVelEpsEff THEN
            eState := E_DL_StopState.eSettling; // 速度已跌到阈值以下，进稳定确认 / the speed fell below the threshold, settle
        END_IF
    E_DL_StopState.eSettling :
        bBusy := TRUE;                         // 稳定确认中仍算忙 / settling still counts as busy
        uState := DL_STOP_UI_SETTLE;           // 状态镜像 / state mirror
        IF fbSettle.Q THEN
            eState := E_DL_StopState.eDone;    // 稳定窗到期即完成 / the settle window expiring completes the stop
            bDone := TRUE;                     // 完成单拍脉冲 / the single-cycle done pulse
            bStopped := TRUE;                  // 已静止标志 / the stopped flag
            bBusy := FALSE;                    // 完成后不忙 / no longer busy after completion
        END_IF
    E_DL_StopState.eDone :
        bBusy := FALSE;                        // 完成态不忙 / the done state is not busy
        bStopped := TRUE;                      // 保持静止标志 / keep the stopped flag
        uState := DL_STOP_UI_DONE;             // 状态镜像 / state mirror
    E_DL_StopState.eFault :
        bBusy := FALSE;                        // 故障态不忙 / the fault state is not busy
        bStopped := FALSE;                     // 故障态不宣称静止 / the fault state never claims a standstill
        uState := DL_STOP_UI_FAULT;            // 状态镜像 / state mirror
ELSE
    eState := E_DL_StopState.eFault;           // 非法状态一律回安全故障态 / any illegal state falls back to the safe fault state
    eErr := 16#0004_02DA;                      // 本件专用兜底码，用途固定不得改作他用 / the dedicated fallback code, its purpose is fixed
    bError := TRUE;                            // 置故障标志 / raise the error flag
    bBusy := FALSE;                            // 清忙标志 / clear the busy flag
    bStopped := FALSE;                         // 清静止标志 / clear the stopped flag
    uState := DL_STOP_UI_FAULT;                // 状态镜像 / state mirror
END_CASE
END_FUNCTION_BLOCK

(* ---- FB_DL_AxisTeachOffset.st ---- *)
(*==============================================================================
 * 组件名称 (Component)  : FB_DL_AxisTeachOffset
 * 所属子库 (Sublibrary) : DL_Motion
 * 当前版本 (Version)    : 1.0.0
 * 兼容性   (Platform)   : CODESYS 3.5+ / TwinCAT 3 / 汇川 InoProShop / 施耐德 Machine Expert
 *                         仅依赖 Standard.library（R_TRIG），零厂商私有库
 * 功能描述 (Function)   : 示教点与配方偏移管理。① 示教：bTeach 上升沿在轴静止（外部注入
 *                         bAxisStandstill 为真）时把当前 fPosAct 锁存进 _fTaughtPos；运动中
 *                         示教一律拒绝并置信息级（防采样到抖动位置，这是现场示教偏移的
 *                         首要误差源）；② 应用偏移：bApplyOffset 上升沿把 fOffsetValue 写入
 *                         配方偏移槽，写入前先算候选目标位（示教位 + 偏移）并做软限校验，
 *                         **越限则拒绝且原偏移保持不被覆盖**（先判后写，绝不先写后判）。
 * 接口     (Interface)  : 输入 fPosAct 当前实际位置、bTeach 示教命令、bApplyOffset 应用偏移命令、
 *                         fOffsetValue 待写入偏移值、fSoftLo / fSoftHi 轴软限、bAxisStandstill
 *                         外部注入的静止位、bReset 复位；输出 fTaughtPos 已示教位置、fOffsetApplied
 *                         当前生效偏移、bTeachOk 示教受理成功单拍位、eState / eCause / bError / nErrId。
 * 边界     (Boundary)   : ① 组态闸：fSoftHi <= fSoftLo 或任一浮点引脚 NaN → 故障锁存；
 *                         ② 越软限拦截按「候选目标位 = 示教位 + 待写入偏移」判定，判定通过后才
 *                         写偏移槽（写点唯一，无先写后判路径）；
 *                         ③ 非有限位置 → 故障闸，示教不受理（不把 NaN 写进示教槽，R133）；
 *                         ④ R_TRIG 三枚（示教/应用/复位）段 0 无条件周期刷新；
 *                         ⑤ 故障相迁出唯一路径 = bReset 上升沿；⑥ 零全局耦合（无 GVL / 无物理地址）。
 * 分工声明 (Scope)      : 本件只管理示教值与配方偏移，**不下发定位指令、不判断轴是否到位**；
 *                         轴状态与运动指令唯一属主为 `I_DL_MotionAxis`。
 * 解除式   (Release)    : bReset 上升沿 ∧ 组态合法 ∧ 越限条件已解除（当拍候选目标位落在
 *                         〔fSoftLo, fSoftHi〕内，全为当拍量，R240 范式）。
 *                         自证可满足（终审两式 1）：解除式只含当拍比较，偏移值或示教位修正后
 *                         即可达；不含计时器输出与锁存量比较，无恒假因子。
 * 码表     (Codes)      : 16#0004_03B6 故障级：示教偏移故障总码（组态非法 / 目标位越软限 /
 *                         非法相位），锁存至 bReset 上升沿，归因由 eCause 承载（R190 单件单总码）；
 *                         16#0004_04B6 信息级：运动中示教被拒绝（信息级，不锁故障）。
 *                         加码反证（R90）：拒绝示教时 fTaughtPos 保持旧值、bTeachOk 为假，
 *                         该否决若不留码则 HMI 上「操作员按了示教但没生效」完全不可观测
 *                         （bTeachOk 是单拍位且为假），故立一码。
 *                         码段说明：0004 段故障子带 03xx / 信息子带 04xx，本件取 03B6 / 04B6
 *                         （源码实扫该两槽为空，续接同子带已用最大值，未回填碎片孔洞）。
 * 开源溯源 (Origin)     : 道莅自研 clean-room（参考示教-配方偏移现场惯例与参数域，零代码行复制；
 *                         t1-6-plcopen 族）
 * 修订历史 (Revision)   : 2026-11-19  v1.0.0  R45 首版（批次 3 · 序号 12）
 *==============================================================================*)

TYPE E_DL_AtoState :
(
    eIdle  := 0,     // 未示教（无有效示教值） / Idle, no valid taught position yet
    eRun   := 10,    // 示教值就绪，可应用偏移 / Taught value ready, offset applicable
    eFault := 90     // 故障锁存相 / Fault latched phase
);
END_TYPE

TYPE E_DL_AtoCause :
(
    eNone       := 0,   // 无故障成因 / No cause
    eCfgIllegal := 1,   // 组态非法 / Illegal configuration
    eSoftLimit  := 2,   // 候选目标位越软限 / Candidate target outside soft limits
    eNonFinite  := 3,   // 位置或偏移非有限 / Non-finite position or offset
    ePhaseBad   := 4    // 非法相位兜底 / Illegal phase fallback
);
END_TYPE

FUNCTION_BLOCK FB_DL_AxisTeachOffset
VAR_INPUT
    fPosAct        : REAL := 0.0;         // 当前实际位置 [mm] / Current actual position [mm]
    bTeach         : BOOL := FALSE;       // 示教命令，上升沿受理一次 [-] / Teach command, rising edge accepts once
    bApplyOffset   : BOOL := FALSE;       // 应用偏移命令，上升沿受理一次 [-] / Apply-offset command, rising edge accepts once
    fOffsetValue   : REAL := 0.0;         // 待写入的偏移值 [mm] / Offset value to be written [mm]
    fSoftLo        : REAL := -100.0;      // 轴软限下限，域 < fSoftHi [mm] / Soft limit lower bound, domain < fSoftHi [mm]
    fSoftHi        : REAL := 100.0;       // 轴软限上限，域 > fSoftLo [mm] / Soft limit upper bound, domain > fSoftLo [mm]
    bAxisStandstill: BOOL := FALSE;       // 轴静止位（外部注入，示教受理前置） [-] / Axis standstill flag, injected
    bReset         : BOOL := FALSE;       // 复位命令，上升沿清故障 [-] / Reset command, rising edge clears fault
END_VAR
VAR_OUTPUT
    fTaughtPos     : REAL;                // 已示教位置（锁存量回放） [mm] / Taught position, latched replay [mm]
    fOffsetApplied : REAL;                // 当前生效偏移（锁存量回放） [mm] / Effective offset, latched replay [mm]
    bTeachOk       : BOOL;                // 示教受理成功单拍位 [-] / Teach accepted, single scan
    eState         : E_DL_AtoState;       // 状态出口，段 6 单点映射 / State outlet
    eCause         : E_DL_AtoCause;       // 故障成因出口（R190 归因唯一） / Fault cause outlet
    bError         : BOOL;                // 故障锁存标志 [-] / Fault latch flag
    nErrId         : UDINT;               // 事件码，0 = 无事件 / Event code, 0 = no event
END_VAR
VAR
    _eState        : E_DL_AtoState := E_DL_AtoState.eIdle;    // 内部相位（CASE 唯一写入目标） / Internal phase
    _eCause        : E_DL_AtoCause := E_DL_AtoCause.eNone;    // 故障成因锁存（锁存量） / Latched cause
    rtTeach        : R_TRIG;              // 示教沿实例，段 0 无条件调用 / Teach rising edge
    rtApply        : R_TRIG;              // 应用沿实例，段 0 无条件调用 / Apply rising edge
    rtReset        : R_TRIG;              // 复位沿实例，段 0 无条件调用 / Reset edge
    _fTaughtPos    : REAL;                // 示教位置槽（锁存量） [mm] / Taught position slot, latched
    _fOffsetSlot   : REAL;                // 配方偏移槽（锁存量，唯一写入点） [mm] / Recipe offset slot, single write point
    _bTaughtValid  : BOOL;                // 示教槽有效标记（锁存量） [-] / Taught slot valid flag
    _fCand        : REAL;                 // 候选目标位 = 示教位 + 待写入偏移 [mm] / Candidate target, taught plus offset [mm]
    _bNonFin       : BOOL;                // 输入非有限当拍量 [-] / Non-finite input this scan
    _bCfgBad       : BOOL;                // 组态非法当拍量 [-] / Illegal configuration
    _bCandInRange  : BOOL;                // 候选目标位在软限内当拍量 [-] / Candidate target inside soft limits
    _bFault        : BOOL;                // 故障锁存位（锁存量） / Latched fault bit
    _uFault        : UDINT;               // 故障码锁存（锁存量） / Latched fault code
    _uInfo         : UDINT;               // 信息码，每拍重算 / Info code, recomputed each scan
END_VAR
VAR CONSTANT
    DL_FLOAT_EPS : REAL := 1.0E-6;        // 浮点判零容差（软限比较统一口径） [mm] / Float epsilon for zero tests [mm]
END_VAR

(* —— 段 0：当拍判据派生 + 沿实例无条件周期刷新 —— *)
_bNonFin := (fPosAct <> fPosAct) OR (fOffsetValue <> fOffsetValue)                        // NaN 自反判（判等禁令唯一例外） / NaN self-reflexive tests
          OR (fSoftLo <> fSoftLo) OR (fSoftHi <> fSoftHi)                                // 软限 NaN 判 / Soft limit NaN tests
          OR ((fPosAct - fPosAct) <> (fPosAct - fPosAct))                                // 位置 Inf 差值自减判 / Inf test on position
          OR ((fOffsetValue - fOffsetValue) <> (fOffsetValue - fOffsetValue));            // 偏移 Inf 差值自减判 / Inf test on offset
_bCfgBad := (fSoftHi <= fSoftLo) OR ((fSoftHi - fSoftLo) <= DL_FLOAT_EPS);                // 软限几何组态闸（R151） / Soft-limit geometry gate
_fCand  := _fTaughtPos + fOffsetValue;                                                   // 候选目标位 / Candidate target position
_bCandInRange := (_fCand >= fSoftLo) AND (_fCand <= fSoftHi);                             // 候选位在软限内当拍量 / Candidate inside soft limits
rtTeach(CLK := bTeach);                                                                   // 示教沿，每拍必调（R228A） / Teach edge, called every scan
rtApply(CLK := bApplyOffset);                                                             // 应用沿，每拍必调 / Apply edge, called every scan
rtReset(CLK := bReset);                                                                   // 复位沿，每拍必调 / Reset edge, called every scan

(* —— 段 1：单拍量预清零（锁存量不入清单，R107） —— *)
_uInfo         := 16#0000_0000;        // 信息码每拍重算 / Info recomputed every scan
bTeachOk       := FALSE;               // 示教成功位每拍预清，唯一分支置位（R44 范式） / Teach-ok preset
nErrId         := 16#0000_0000;        // 事件码缺省无事件 / Event code default none
bError         := FALSE;               // 故障标志每拍预清，故障分支同拍置位（R45 配对） / Flag preset

(* —— 段 2：复位沿 + 组态域闸 + 非有限闸 —— *)
IF rtReset.Q THEN                                                        // 当拍复位沿 / current-scan reset edge
    _bFault := FALSE;                                                    // 清故障锁存位（锁存量） / Clear fault latch
    _uFault := 16#0000_0000;                                             // 清故障锁存码（锁存量） / Clear latched code
    _eCause := E_DL_AtoCause.eNone;                                      // 清成因（锁存量） / Clear latched cause
    IF _eState = E_DL_AtoState.eFault THEN
        _eState := E_DL_AtoState.eIdle;                                  // 故障相迁出唯一路径 / Sole exit from fault phase
    END_IF
END_IF
IF _bCfgBad THEN                                                         // 组态域闸 / Configuration gate
    _uFault := 16#0004_03B6;                                             // 故障级：示教偏移故障总码 / Fault-level: teach/offset fault code
    _bFault := TRUE;
    bError  := TRUE;                                                     // 故障标志同拍置位（R45 配对） / Error flag set same scan
    _eCause := E_DL_AtoCause.eCfgIllegal;                                // 归因：组态非法 / Cause: illegal configuration
END_IF
IF (NOT _bFault) AND _bNonFin THEN                                       // 位置/偏移非有限 / Non-finite position or offset
    _uFault := 16#0004_03B6;
    _bFault := TRUE;
    bError  := TRUE;
    _eCause := E_DL_AtoCause.eNonFinite;                                 // 归因：非有限 / Cause: non-finite
END_IF

(* —— 段 3：示教授理（静止前置 + 非有限拒收） —— *)
IF (NOT _bFault) AND rtTeach.Q THEN                                      // 示教上升沿（当拍量） / Teach rising edge
    IF bAxisStandstill THEN                                              // 静止前置满足才受理 / Accept only at standstill
        _fTaughtPos := fPosAct;                                          // 锁存当前位置（示教槽唯一写入点） / Latch current position
        _bTaughtValid := TRUE;                                           // 示教槽置有效 / Mark taught slot valid
        bTeachOk := TRUE;                                                // 单拍成功位 / Single-scan success flag
    ELSE
        _uInfo := 16#0004_04B6;                                          // 信息级：运动中示教被拒绝 / Info: teach rejected while moving
    END_IF
END_IF

(* —— 段 4：应用偏移（先判软限后写槽，绝不先写后判） —— *)
IF (NOT _bFault) AND rtApply.Q THEN                                      // 应用上升沿（当拍量） / Apply rising edge
    IF _bTaughtValid AND _bCandInRange THEN                              // 前置齐备且候选位在软限内 / Preconditions met and candidate in range
        _fOffsetSlot := fOffsetValue;                                    // 写偏移槽（唯一写入点，判定通过后才写） / Write offset slot only after the check passes
    ELSE
        _uFault := 16#0004_03B6;                                         // 故障级：候选目标位越软限（或未示教） / Fault-level: candidate outside limits or not taught
        _bFault := TRUE;
        bError  := TRUE;                                                 // 故障标志同拍置位（R45 配对） / Error flag set same scan
        _eCause := E_DL_AtoCause.eSoftLimit;                             // 归因：越软限 / Cause: soft limit
    END_IF
END_IF

(* —— 段 5：故障解除式（R240 全当拍量） —— *)
IF rtReset.Q AND (NOT _bCfgBad) AND (NOT _bNonFin) AND (_bCandInRange OR (NOT _bTaughtValid)) THEN
    _bFault := FALSE;                                                    // 清故障锁存位（锁存量） / Clear fault latch
    _uFault := 16#0000_0000;                                             // 清故障锁存码（锁存量） / Clear latched code
    _eCause := E_DL_AtoCause.eNone;                                      // 清成因（锁存量） / Clear latched cause
END_IF

(* —— 段 5A：故障锁存相位迁移闸 —— *)
IF _bFault AND (_eState <> E_DL_AtoState.eFault) THEN
    _eState := E_DL_AtoState.eFault;                                     // 锁存即入故障相 / Latch enters fault phase
END_IF

(* —— 段 6：相位机（ENUM 全成员显式标签 + ELSE 兜底，R128） —— *)
CASE _eState OF

E_DL_AtoState.eIdle:
    IF _bTaughtValid AND (NOT _bFault) THEN                              // 出口 1：示教槽已就绪 / Taught slot ready
        _eState := E_DL_AtoState.eRun;
    ELSIF _bFault THEN                                                   // 出口 2：故障锁存 / Fault latched
        _eState := E_DL_AtoState.eFault;
    END_IF

E_DL_AtoState.eRun:
    IF (NOT _bTaughtValid) THEN                                          // 出口 1：示教槽失效（前置消失，R98） / Taught slot invalid
        _eState := E_DL_AtoState.eIdle;
    ELSIF _bFault THEN                                                   // 出口 2：故障锁存 / Fault latched
        _eState := E_DL_AtoState.eFault;
    END_IF

E_DL_AtoState.eFault:
    ;                                                                     // 故障相：仅段 5 复位沿可迁出 / Only the reset edge leaves this phase

ELSE
    _uFault := 16#0004_03B6;                                             // 故障级：非法相位兜底（归并总码） / Illegal-phase fallback
    _bFault := TRUE;
    bError  := TRUE;
    _eCause := E_DL_AtoCause.ePhaseBad;                                  // 归因：非法相位 / Cause: illegal phase
    _eState := E_DL_AtoState.eFault;

END_CASE

(* —— 段 7：出口单点映射（名实同源；锁存码回放） —— *)
fTaughtPos     := _fTaughtPos;                                           // 示教位出口（锁存量回放） / Taught position outlet
fOffsetApplied := _fOffsetSlot;                                          // 生效偏移出口（锁存量回放） / Effective offset outlet
IF _bFault THEN
    bTeachOk := FALSE;                                                   // 故障相不宣称示教成功 / No success claim in fault
    nErrId   := _uFault;                                                 // 故障锁存码回放 / Replay latched fault code
ELSE
    nErrId   := _uInfo;                                                  // 信息码 / Info code
END_IF
bError := _bFault;                                                       // 故障标志与锁存同源（名实双出口，R191） / Flag from latch
eState := _eState;                                                       // 状态出口 / State outlet
eCause := _eCause;                                                       // 成因出口 / Cause outlet

END_FUNCTION_BLOCK

(* ---- FB_DL_AxisThermalComp.st ---- *)
(*==============================================================================
 * 组件名称 (Component)  : FB_DL_AxisThermalComp
 * 所属子库 (Sublibrary) : DL_Motion
 * 当前版本 (Version)    : 1.0.0
 * 兼容性   (Platform)   : CODESYS 3.5+ / TwinCAT 3 / 汇川 InoProShop / 施耐德 Machine Expert
 *                         仅依赖 Standard.library（ABS），零厂商私有库
 * 功能描述 (Function)   : 轴热变形行程比例补偿：温度差 fTempDiffK（相对参考温，
 *                         K）经一阶热模型（时间常数 fTauS 可配）滤波后乘热
 *                         膨胀标度 fScaleUmK（µm/K）换算为行程补偿量：
 *                           α = fCy ÷ (fTauS + fCy)（离散一阶步长，域钳 [0,1]）
 *                           fFiltK = fFiltK + α × (fTempDiffK − fFiltK)
 *                           fCompValMm = fFiltK × fScaleUmK ÷ 1000
 *                         温度超域（|fTempDiffK| > fTMaxK）钳位并置信息码
 *                         eTempClamped；bEnable=FALSE 直通输出 0（规格指定，
 *                         R191 声明：未使能期强制归零而非冻结保持）。
 * 接口     (Interface)  : 输入 fTempDiffK 温度差（相对参考温） [K]、fScaleUmK
 *                         热膨胀标度（域 > 0） [µm/K]、fTauS 一阶热模型时间
 *                         常数（域 > 0） [s]、fTMaxK 温度差域半宽（域 > 0）
 *                         [K]、fCycle 扫描周期（<=0 用缺省） [s]、bEnable
 *                         使能、bReset 复位；输出 fCompValMm 行程补偿
 *                         [mm]、fFiltK 滤波后温度差（诊断透读） [K]、
 *                         eErrCode 错误码、bError 故障标志。
 * 边界     (Boundary)   : ① **属主边界（写死）：本件只算热补偿量，不测温度、
 *                         不接管轴使能**；温度采集归模拟量输入层。
 *                         ② 步长 α：fTauS <= 0 走组态锁存（规格域 > 0），
 *                         正常域 α = fCy/(fTauS+fCy) ∈ (0,1) 结构性稳定
 *                         （分母两项恒正，无除零）。
 *                         ③ 非有限判据（R79 双判）先行：温度差/标度非有限时
 *                         输出保持上次滤波值对应补偿量（冻结），置信息码
 *                         eInputHold，不污染滤波态。
 *                         ④ 组态闸：fScaleUmK <= 0、fTauS <= 0、fTMaxK <= 0
 *                         → 锁存故障，输出强制 0，解除沿 = bReset 上升沿。
 *                         ⑤ µm→mm 换算用常量除法（÷1000 非零常量，无除零）。
 *                         ⑥ 零全局耦合（无 GVL / VAR_EXTERNAL / 物理地址）。
 * 分工声明 (Scope)      : 与 `FB_DL_AxisScrewPitchComp` 分工：几何螺距误差归
 *                         那件、热变形比例项归本件；与 `FB_DL_LeadLagCompensator`
 *                         分工：通用超前滞后归那件，本件内嵌一阶滤波为热模型
 *                         属主实现（不引用，独立验收）。
 * 来源标签 (Source Tag) : 自研线（一阶热模型与线性热膨胀为公开物理定义 clean-room）
 * 码表     (Codes)      : 本件不占用任何全局数字码位。出口为 LREAL 组 +
 *                         ENUM 错误码；数字码位待主控收口阶段统一派号。
 * 红线自检 (Redline)    : R1 ✓ 零 GVL/VAR_EXTERNAL ｜ R2 ✓ 零 %I/%Q/%M ｜ R3 ✓ 纯 IEC 61131-3
 *                         R4 ✓ 步长域稳定 + 温度域钳位 + 非有限冻结 + 组态锁存
 *                         ｜ R5 ✓ 声明逐行同行双语注释
 *                         R6 N/A（无 ENUM 状态机） ｜ R7 ✓ 一 R_TRIG 段 0 无条件刷新
 * 修订历史 (Revision)   : 2026-11-20  v1.0.0  R50 首版（批次 2 · 序号 8）
 * 验收向量 (Acceptance) : ① fScaleUmK=10, fTauS=60, fCycle=0.01：温度差恒
 *                         20 K 滤波收敛后 fFiltK→20，fCompValMm = 20×10÷1000
 *                         = 0.2 mm（稳态，eOk）；② 温度差 100 K，fTMaxK=80
 *                         → 钳 80 → 收敛后 fCompValMm = 0.8 mm，
 *                         eTempClamped；③ bEnable=FALSE → fCompValMm=0
 *                         （直通零，规格声明）；④ fTauS=0 → 锁存 eCfgBad。
 *==============================================================================*)

(*-----------------------------------------------------------------------------
 * 枚举: E_DL_AtcErr（错误码；信息级不置 bError，故障级恒伴 bError=TRUE）
 *----------------------------------------------------------------------------*)
TYPE E_DL_AtcErr :
(
    eOk          := 0,   // 正常 / Normal
    eCfgBad      := 1,   // 故障级：组态非法（标度/时间常数/域半宽） / Fault: illegal configuration
    eTempClamped := 2,   // 信息级：温度差超域已钳位 / Info: temperature diff clamped
    eInputHold   := 3    // 信息级：输入非有限，滤波态冻结 / Info: non-finite input, filter state frozen
);
END_TYPE

FUNCTION_BLOCK FB_DL_AxisThermalComp
VAR_INPUT
    fTempDiffK : LREAL := 0.0;        // 温度差（相对参考温） [K] / Temperature difference from reference [K]
    fScaleUmK  : LREAL := 10.0;       // 热膨胀标度，域 > 0 [µm/K] / Thermal expansion scale [um/K]
    fTauS      : LREAL := 60.0;       // 一阶热模型时间常数，域 > 0 [s] / First-order thermal time constant [s]
    fTMaxK     : LREAL := 80.0;       // 温度差域半宽（对称 ±），域 > 0 [K] / Temperature domain half-width [K]
    fCycle     : LREAL := 0.0;        // 扫描周期（<=0 用缺省） [s] / Scan cycle, default used when <= 0
    bEnable    : BOOL := FALSE;       // 使能（FALSE=输出直通 0，规格声明） [-] / Enable, FALSE forces zero output
    bReset     : BOOL := FALSE;       // 复位，上升沿清组态故障锁存 [-] / Reset, rising edge clears cfg latch
END_VAR
VAR_OUTPUT
    fCompValMm : LREAL;               // 行程补偿输出（叠加位置设定侧） [mm] / Travel compensation output [mm]
    fFiltK     : LREAL;               // 滤波后温度差（诊断透读） [K] / Filtered temperature difference [K]
    eErrCode   : E_DL_AtcErr;         // 错误码出口 / Error code outlet
    bError     : BOOL;                // 故障标志（组态锁存） [-] / Error flag, latched
END_VAR
VAR
    _fFilt    : LREAL := 0.0;         // 滤波温度差锁存（冻结源） [K] / Filtered temperature latch
    _fCy      : LREAL;                // 当拍有效周期 [s] / Effective cycle this scan
    _fAlpha   : LREAL;                // 离散一阶步长（域 (0,1)） [-] / Discrete first-order step
    _fTempUse : LREAL;                // 钳位后温度差 [K] / Clamped temperature difference
    _bNonFin  : BOOL;                 // 输入非有限当拍量 [-] / Non-finite input this scan
    _bClamped : BOOL;                 // 本拍发生温度钳位 [-] / Temperature clamped this scan
    _bCfgBad  : BOOL;                 // 组态非法当拍量 [-] / Illegal configuration this scan
    _bErrLatch: BOOL;                 // 组态故障锁存位（解除沿 = bReset 上升沿） / Latched config fault
    rtReset   : R_TRIG;               // 复位沿实例，段 0 无条件调用 / Reset edge instance
END_VAR
VAR CONSTANT
    DL_ATC_CYDEF  : LREAL := 0.01;    // 缺省扫描周期 [s] / Default scan cycle
    DL_ATC_UM2MM  : LREAL := 1000.0;  // µm→mm 换算常量（非零，无除零） [µm/mm] / um per mm constant
    DL_ATC_ZERO   : LREAL := 0.0;     // 判零基准 [K] / Zero base
    DL_ATC_ONE    : LREAL := 1.0;     // 步长钳位上界 [-] / Step ceiling
END_VAR

(* —— 段 0：非有限判 + 组态闸 + 周期派生 + 沿刷新 —— *)
_bNonFin := (fTempDiffK <> fTempDiffK) OR ((fTempDiffK - fTempDiffK) <> DL_ATC_ZERO)
         OR (fScaleUmK <> fScaleUmK) OR ((fScaleUmK - fScaleUmK) <> DL_ATC_ZERO);   // 输入非有限（R79 双判） / Non-finite inputs
_bCfgBad := (fScaleUmK <= DL_ATC_ZERO) OR (fTauS <= DL_ATC_ZERO) OR (fTMaxK <= DL_ATC_ZERO);   // 组态域闸 / Configuration gate
IF fCycle > DL_ATC_ZERO THEN
    _fCy := fCycle;                                // 组态周期有效 / Configured cycle valid
ELSE
    _fCy := DL_ATC_CYDEF;                          // 周期缺省兜底 / Default cycle fallback
END_IF
rtReset(CLK := bReset);                            // 复位沿，每拍必调 / Reset edge, every scan

(* —— 段 1：复位沿与组态锁存 —— *)
IF rtReset.Q THEN
    _bErrLatch := FALSE;                           // 清组态锁存（R188 声明：解除沿 = bReset 上升沿） / Clear cfg latch
END_IF
IF _bCfgBad AND (NOT _bErrLatch) THEN
    _bErrLatch := TRUE;                            // 锁存 / Latch
END_IF

(* —— 段 2：温度域钳位（非有限冻结滤波态，不污染） —— *)
_bClamped := FALSE;                                // 钳位量预清 / Clamp preset
_fTempUse := DL_ATC_ZERO;                          // 安全侧起步 0 / Safe-side start
IF (NOT _bErrLatch) AND (NOT _bNonFin) THEN
    _fTempUse := fTempDiffK;                       // 温度差工作副本 / Temperature working copy
    IF _fTempUse > fTMaxK THEN
        _fTempUse := fTMaxK;                       // 超上域钳位（规格） / Clamp high
        _bClamped := TRUE;                         // 记钳位 / Mark clamp
    ELSIF _fTempUse < (-fTMaxK) THEN
        _fTempUse := -fTMaxK;                      // 超下域钳位（对称 ±） / Clamp low symmetric
        _bClamped := TRUE;                         // 记钳位 / Mark clamp
    END_IF
END_IF

(* —— 段 3：一阶热模型递推与补偿合成（故障期冻结；未使能直通 0） —— *)
IF (NOT _bErrLatch) AND (NOT _bNonFin) THEN
    _fAlpha := _fCy / (fTauS + _fCy);              // 步长（分母两项恒正，无除零；fTauS>0 已闸） / Step size
    _fFilt := _fFilt + _fAlpha * (_fTempUse - _fFilt);   // 一阶热模型递推 / First-order thermal recursion
    IF bEnable THEN
        fCompValMm := _fFilt * fScaleUmK / DL_ATC_UM2MM;   // 补偿 = 滤波温差×标度÷1000 [mm] / Compensation synthesis
    ELSE
        fCompValMm := DL_ATC_ZERO;                 // 未使能直通 0（R191 声明：强制归零） / Disabled: forced zero
    END_IF
ELSIF (NOT _bErrLatch) AND _bNonFin THEN
    fCompValMm := _fFilt * fScaleUmK / DL_ATC_UM2MM;   // 非有限冻结：按上次滤波值输出（头注释③） / Freeze at last filtered value
ELSE
    fCompValMm := DL_ATC_ZERO;                     // 故障安全侧 0 / Fault safe-side zero
END_IF

(* —— 段 4：出口单点映射（名实双出口同源，R191） —— *)
fFiltK := _fFilt;                                  // 滤波温差透读出口 / Filtered temperature readout
IF _bErrLatch THEN
    bError := TRUE;                                // 故障标志（R45 配对） / Error flag
    eErrCode := E_DL_AtcErr.eCfgBad;               // 故障级码 / Fault code
ELSE
    bError := FALSE;                               // 无故障级条件 / No fault
    IF _bNonFin THEN
        eErrCode := E_DL_AtcErr.eInputHold;        // 信息级：冻结口径 / Info: frozen
    ELSIF _bClamped THEN
        eErrCode := E_DL_AtcErr.eTempClamped;      // 信息级：钳位口径 / Info: clamped
    ELSE
        eErrCode := E_DL_AtcErr.eOk;               // 正常 / Normal
    END_IF
END_IF

END_FUNCTION_BLOCK

(* ---- FB_DL_AxisTorqueFeedforward.st ---- *)
(*==============================================================================
 * 组件名称 (Component)  : FB_DL_AxisTorqueFeedforward
 * 所属子库 (Sublibrary) : DL_Motion
 * 当前版本 (Version)    : 1.0.0
 * 兼容性   (Platform)   : CODESYS 3.5+ / TwinCAT 3 / 汇川 InoProShop / 施耐德 Machine Expert
 *                         仅依赖 Standard.library（ABS），零厂商私有库
 * 功能描述 (Function)   : 转矩前馈合成（刚体动力学 + 黏性摩擦项）：
 *                           fTorqueFF = fJ × fAccel + fVisc × fVel
 *                         输出限幅 ±fMax（必填，域 > 0，超限钳位并置信息码
 *                         eClamped）；J <= 0 → 拒算直通 0 并置信息码 eJInvalid
 *                         （规格指定）；非有限输入 → 输出 0、信息码 eInputHold。
 * 接口     (Interface)  : 输入 fAccel 角加速度 [rad/s²]、fJ 转动惯量（域 > 0
 *                         参算，<=0 拒算） [kg·m²]、fVisc 黏性摩擦系数
 *                         [N·m·s/rad]、fVel 角速度 [rad/s]、fMax 输出限幅
 *                         （必填，域 > 0） [N·m]、bReset 复位；输出 fTorqueFF
 *                         转矩前馈 [N·m]、eErrCode 错误码、bError 故障标志。
 * 边界     (Boundary)   : ① **属主边界（写死）：本件只算前馈标量，不做摩擦
 *                         辨识、不接管轴使能**；辨识归 `FB_DL_AxisInertiaIdent`
 *                         / `FB_DL_AxisFrictionFf`。
 *                         ② J <= 0 拒算直通 0（规格指定，物理上负/零惯量
 *                         无刚体动力学意义）；fVisc/fVel 不参与拒算域闸
 *                         （黏性项可独立为零）。
 *                         ③ fMax 必填闸：fMax <= 0 或非有限 → 锁存故障
 *                         eCfgBad，输出 0（限幅缺失时钳位语义不成立，不得
 *                         放行无界前馈），解除沿 = bReset 上升沿（R45 配对）。
 *                         ④ 非有限判据（R79 双判）：四个动力学量逐一双判；
 *                         拒算/非有限输出 0 均为信息级（不置 bError）。
 *                         ⑤ 限幅对称 ±fMax，钳位后信息码 eClamped（信息级）。
 *                         ⑥ 零全局耦合（无 GVL / VAR_EXTERNAL / 物理地址）。
 * 分工声明 (Scope)      : 与 `FB_DL_AxisFrictionFf` 分工：摩擦辨识与库仑项归
 *                         那件，本件黏性项为线性合成（系数直传）；与
 *                         `FB_DL_AxisCoggingFf` 分工：齿槽补偿归那件。
 * 来源标签 (Source Tag) : 自研线（刚体动力学 τ=Jα+Bω 为公开物理定义 clean-room）
 * 码表     (Codes)      : 本件不占用任何全局数字码位。出口为 LREAL 转矩 +
 *                         ENUM 错误码；数字码位待主控收口阶段统一派号。
 * 红线自检 (Redline)    : R1 ✓ 零 GVL/VAR_EXTERNAL ｜ R2 ✓ 零 %I/%Q/%M ｜ R3 ✓ 纯 IEC 61131-3
 *                         R4 ✓ J 域拒算 + fMax 必填锁存 + 非有限双判 + 限幅
 *                         ｜ R5 ✓ 声明逐行同行双语注释
 *                         R6 N/A（无 ENUM 状态机） ｜ R7 ✓ 一 R_TRIG 段 0 无条件刷新
 * 修订历史 (Revision)   : 2026-11-20  v1.0.0  R50 首版（批次 3 · 序号 15）
 * 验收向量 (Acceptance) : ① fJ=0.01, fAccel=100, fVisc=0.005, fVel=1000,
 *                         fMax=10 → 0.01×100 + 0.005×1000 = 1.0 + 5.0 =
 *                         6.0 N·m，eOk；② 同输入 fMax=5 → 钳 ±5 → 5.0 N·m，
 *                         eClamped；③ fJ=0 → 输出 0，eJInvalid（fVisc×fVel
 *                         项一并拒算，规格①口径）；④ fMax=0 → 锁存 eCfgBad，
 *                         输出 0。
 *==============================================================================*)

(*-----------------------------------------------------------------------------
 * 枚举: E_DL_TffErr（错误码；信息级不置 bError，故障级恒伴 bError=TRUE）
 *----------------------------------------------------------------------------*)
TYPE E_DL_TffErr :
(
    eOk        := 0,   // 正常 / Normal
    eCfgBad    := 1,   // 故障级：fMax 必填闸破约（<=0 或非有限） / Fault: fMax mandatory gate violated
    eClamped   := 2,   // 信息级：输出超 ±fMax 已钳位 / Info: output clamped
    eJInvalid  := 3,   // 信息级：J<=0 拒算直通 0 / Info: non-positive J, zero output
    eInputHold := 4    // 信息级：动力学量非有限，输出 0 / Info: non-finite input, zero output
);
END_TYPE

FUNCTION_BLOCK FB_DL_AxisTorqueFeedforward
VAR_INPUT
    fAccel : LREAL := 0.0;            // 角加速度 [rad/s2] / Angular acceleration
    fJ     : LREAL := 0.01;           // 转动惯量（<=0 拒算） [kg·m2] / Inertia, non-positive rejects
    fVisc  : LREAL := 0.005;          // 黏性摩擦系数 [N·m·s/rad] / Viscous friction coefficient
    fVel   : LREAL := 0.0;            // 角速度 [rad/s] / Angular velocity
    fMax   : LREAL := 10.0;           // 输出限幅（必填，对称 ±），域 > 0 [N·m] / Torque limit, mandatory
    bReset : BOOL := FALSE;           // 复位，上升沿清组态故障锁存 [-] / Reset, rising edge clears cfg latch
END_VAR
VAR_OUTPUT
    fTorqueFF : LREAL;                // 转矩前馈输出（已限幅） [N·m] / Torque feedforward output
    eErrCode  : E_DL_TffErr;          // 错误码出口 / Error code outlet
    bError    : BOOL;                 // 故障标志（fMax 必填锁存） [-] / Error flag, latched
END_VAR
VAR
    _fRaw     : LREAL;                // 未限幅合成转矩 [N·m] / Raw composed torque
    _bJBad    : BOOL;                 // J 拒算当拍量 [-] / J rejection this scan
    _bNonFin  : BOOL;                 // 动力学量非有限当拍量 [-] / Non-finite dynamics this scan
    _bClamped : BOOL;                 // 本拍发生限幅 [-] / Clamped this scan
    _bCfgBad  : BOOL;                 // fMax 必填闸破约当拍量 [-] / fMax gate violation
    _bErrLatch: BOOL;                 // 组态故障锁存位（解除沿 = bReset 上升沿） / Latched config fault
    rtReset   : R_TRIG;               // 复位沿实例，段 0 无条件调用 / Reset edge instance
END_VAR
VAR CONSTANT
    DL_TFF_ZERO : LREAL := 0.0;       // 拒算输出与判零基准 [N·m] / Zero output and base
END_VAR

(* —— 段 0：非有限判 + 必填闸 + 沿刷新 —— *)
_bNonFin := (fAccel <> fAccel) OR ((fAccel - fAccel) <> DL_TFF_ZERO)
         OR (fJ <> fJ) OR ((fJ - fJ) <> DL_TFF_ZERO)
         OR (fVisc <> fVisc) OR ((fVisc - fVisc) <> DL_TFF_ZERO)
         OR (fVel <> fVel) OR ((fVel - fVel) <> DL_TFF_ZERO);   // 动力学量非有限（R79 双判） / Non-finite dynamics
_bCfgBad := (fMax <= DL_TFF_ZERO) OR (fMax <> fMax) OR ((fMax - fMax) <> DL_TFF_ZERO);   // fMax 必填闸（域 + 非有限） / fMax mandatory gate
rtReset(CLK := bReset);               // 复位沿，每拍必调 / Reset edge, every scan

(* —— 段 1：复位沿与组态锁存 —— *)
IF rtReset.Q THEN
    _bErrLatch := FALSE;              // 清组态锁存（R188 声明：解除沿 = bReset 上升沿） / Clear cfg latch
END_IF
IF _bCfgBad AND (NOT _bErrLatch) THEN
    _bErrLatch := TRUE;               // 锁存 / Latch
END_IF

(* —— 段 2：拒算判据（J<=0 与非有限并行记录，信息级） —— *)
_bJBad := (fJ <= DL_TFF_ZERO);        // J 拒算判据（规格②） / J rejection test

(* —— 段 3：转矩合成与限幅（故障/J 拒算/非有限 → 输出 0） —— *)
IF _bErrLatch THEN
    fTorqueFF := DL_TFF_ZERO;         // 故障安全侧 0（头注释③） / Fault safe-side zero
ELSIF _bNonFin THEN
    fTorqueFF := DL_TFF_ZERO;         // 非有限输出 0（规格） / Non-finite zero
ELSIF _bJBad THEN
    fTorqueFF := DL_TFF_ZERO;         // J<=0 拒算直通 0（规格②） / J rejection zero
ELSE
    _fRaw := fJ * fAccel + fVisc * fVel;   // 刚体 + 黏性合成 [N·m] / Rigid + viscous synthesis
    _bClamped := FALSE;               // 限幅量预清 / Clamp preset
    IF _fRaw > fMax THEN
        _fRaw := fMax;                // 上限钳位 / Clamp high
        _bClamped := TRUE;            // 记钳位 / Mark clamp
    ELSIF _fRaw < (-fMax) THEN
        _fRaw := -fMax;               // 下限钳位（对称 ±） / Clamp low symmetric
        _bClamped := TRUE;            // 记钳位 / Mark clamp
    END_IF
    fTorqueFF := _fRaw;               // 前馈出口（已限幅） / Feedforward outlet
END_IF

(* —— 段 4：出口单点映射（错误码归约，R191） —— *)
IF _bErrLatch THEN
    bError := TRUE;                   // 故障标志（R45 配对） / Error flag
    eErrCode := E_DL_TffErr.eCfgBad;  // 故障级码 / Fault code
ELSE
    bError := FALSE;                  // 无故障级条件 / No fault
    IF _bNonFin THEN
        eErrCode := E_DL_TffErr.eInputHold;   // 信息级：非有限口径 / Info: non-finite
    ELSIF _bJBad THEN
        eErrCode := E_DL_TffErr.eJInvalid;    // 信息级：J 拒算口径 / Info: J rejected
    ELSIF _bClamped THEN
        eErrCode := E_DL_TffErr.eClamped;     // 信息级：钳位口径 / Info: clamped
    ELSE
        eErrCode := E_DL_TffErr.eOk;          // 正常 / Normal
    END_IF
END_IF

END_FUNCTION_BLOCK
